(* PLC project Codesys Code Execution Speed Tests, CODESYS CODESYS V3.5 SP18 Patch 2, author Toni Kucic *)
(* stored: creationDateTime 2022-11-20T20:47:32.0555446, version 1.0, modificationDateTime 2022-11-20T20:38:51.788641, organization TK Automation *)
(* A collection of programs that measure various execution speeds of code. *)

TYPE dtTestStruct : STRUCT
  dummy1 : USINT := 255;
  Elem1 : INT := -1;
  Id : DWORD := 215215126;
  IdText : STRING := 'Testing for speed';
  dummy2 : ARRAY[0..11] OF DWORD;
  dummy4 : BOOL := FALSE;
  dummy5 : STRING(255) := 'Big array';
  dummy6 : LINT := 1211212723838939;
END_STRUCT;
END_TYPE

TYPE dtBitStruct : STRUCT
  bit1 : BIT;
  bit2 : BIT;
  bit3 : BIT;
  bit4 : BIT;
  bit5 : BIT;
  bit6 : BIT;
  bit7 : BIT;
  bit8 : BIT;
  bit9 : BIT;
  bit10 : BIT;
  bit11 : BIT;
  bit12 : BIT;
  bit13 : BIT;
  bit14 : BIT;
  bit15 : BIT;
  bit16 : BIT;
END_STRUCT;
END_TYPE

TYPE dtSpeedTest : STRUCT
  Results : ARRAY[0..9] OF LTIME;
  Desc : STRING(255);
  AverageExecTime : LTIME;
  OldTime : LTIME;
  ExecTime : LTIME;
END_STRUCT;
END_TYPE

PROGRAM x03_FloatingPointOperations
  VAR CONSTANT
    cNrRuns : USINT(0..9) := 5;
    cRepeatCalcTimes : UDINT := 1000000;  (* 1 Million times *)
  END_VAR
  VAR_INPUT
    vStart : BOOL := FALSE;
  END_VAR
  VAR
    vDone : BOOL := FALSE;
    vRunsCompleted : USINT := 0;
    vStartTime : LTIME;
    vTotalTime : LTIME;
    vTest1 : dtSpeedTest;
    vTest2 : dtSpeedTest;
    vTest3 : dtSpeedTest;
    vTest4 : dtSpeedTest;
    vTest5 : dtSpeedTest;
    vTest6 : dtSpeedTest;
    vTest7 : dtSpeedTest;
    vTest8 : dtSpeedTest;
    vTest9 : dtSpeedTest;
    i : UDINT;
    vInteger1 : INT := 1234;  (* Test vars *)
    vInteger2 : INT := 4231;
    vReal1 : REAL := 1234.4231;
    vReal2 : REAL := 4231.1234;
    vInteger3 : DINT := 1234;
    vInteger4 : DINT := 4231;
    vResult1 : INT;
    vResult2 : REAL;
    vResult3 : DINT;
    vResult4 : INT;
    vResult5 : REAL;
    vResult6 : DINT;
    vResult7 : INT;
    vResult8 : REAL;
    vResult9 : DINT;
  END_VAR

            (*Runs once on event's rising edge*)
vDone 		:= FALSE;
vStartTime 	:= LTIME();

FOR vRunsCompleted:=0 TO cNrRuns DO
	Measure();
END_FOR

vTotalTime := LTIME() - vStartTime;

vTest1.Desc				:= 'Time to add two integers 1 milion times';
vTest1.AverageExecTime 	:= calcAvg(vTest1.Results);
vTest2.Desc				:= 'Time to add two reals 1 milion times';
vTest2.AverageExecTime 	:= calcAvg(vTest2.Results);
vTest3.Desc				:= 'Time to add two DINTs (32b INT) 1 milion times';
vTest3.AverageExecTime 	:= calcAvg(vTest3.Results);
vTest4.Desc				:= 'Time to multiply two integers 1 milion times';
vTest4.AverageExecTime 	:= calcAvg(vTest4.Results);
vTest5.Desc				:= 'Time to multiply two reals 1 milion times';
vTest5.AverageExecTime 	:= calcAvg(vTest5.Results);
vTest6.Desc				:= 'Time to multiply two DINTs (32b INT) 1 milion times';
vTest6.AverageExecTime 	:= calcAvg(vTest6.Results);
vTest7.Desc				:= 'Time to divide two integers 1 milion times';
vTest7.AverageExecTime 	:= calcAvg(vTest7.Results);
vTest8.Desc				:= 'Time to divide two reals 1 milion times';
vTest8.AverageExecTime 	:= calcAvg(vTest8.Results);
vTest9.Desc				:= 'Time to divide two DINTs (32b INT) 1 milion times';
vTest9.AverageExecTime 	:= calcAvg(vTest9.Results);
	
vDone := TRUE;
vStart:= FALSE;

          

ACTION Measure:
                //------------CALCULATION A -------------------
vTest1.OldTime := LTIME();
FOR i:= 0 TO cRepeatCalcTimes DO
	vResult1 := vInteger1 + vInteger2;
END_FOR
vTest1.ExecTime := LTIME() - vTest1.OldTime;

//------------CALCULATION B -------------------
vTest2.OldTime := LTIME();
FOR i:= 0 TO cRepeatCalcTimes DO
	vResult2 := vReal1 + vReal2;
END_FOR
vTest2.ExecTime := LTIME() - vTest2.OldTime;

//------------CALCULATION C -------------------
vTest3.OldTime := LTIME();
FOR i:= 0 TO cRepeatCalcTimes DO
	vResult3 := vInteger3 + vInteger4;
END_FOR
vTest3.ExecTime := LTIME() - vTest3.OldTime;

//------------CALCULATION D -------------------
vTest4.OldTime := LTIME();
FOR i:= 0 TO cRepeatCalcTimes DO
	vResult4 := vInteger1 * vInteger2;
END_FOR
vTest4.ExecTime := LTIME() - vTest4.OldTime;

//------------CALCULATION E -------------------
vTest5.OldTime := LTIME();
FOR i:= 0 TO cRepeatCalcTimes DO
	vResult5 := vReal1 * vReal2;
END_FOR
vTest5.ExecTime := LTIME() - vTest5.OldTime;

//------------CALCULATION F -------------------
vTest6.OldTime := LTIME();
FOR i:= 0 TO cRepeatCalcTimes DO
	vResult6 := vInteger3 * vInteger4;
END_FOR
vTest6.ExecTime := LTIME() - vTest6.OldTime;

//------------CALCULATION G -------------------
vTest7.OldTime := LTIME();
FOR i:= 0 TO cRepeatCalcTimes DO
	vResult7 := vInteger1 / vInteger2;
END_FOR
vTest7.ExecTime := LTIME() - vTest7.OldTime;

//------------CALCULATION H -------------------
vTest8.OldTime := LTIME();
FOR i:= 0 TO cRepeatCalcTimes DO
	vResult8 := vReal1 / vReal2;
END_FOR
vTest8.ExecTime := LTIME() - vTest8.OldTime;

//------------CALCULATION I -------------------
vTest9.OldTime := LTIME();
FOR i:= 0 TO cRepeatCalcTimes DO
	vResult9 := vInteger3 / vInteger4;
END_FOR
vTest9.ExecTime := LTIME() - vTest9.OldTime;


//------------CATCH RESULTS---------------------
vTest1.Results[vRunsCompleted] := vTest1.ExecTime;
vTest2.Results[vRunsCompleted] := vTest2.ExecTime;
vTest3.Results[vRunsCompleted] := vTest3.ExecTime;
vTest4.Results[vRunsCompleted] := vTest4.ExecTime;
vTest5.Results[vRunsCompleted] := vTest5.ExecTime;
vTest6.Results[vRunsCompleted] := vTest6.ExecTime;
vTest7.Results[vRunsCompleted] := vTest7.ExecTime;
vTest8.Results[vRunsCompleted] := vTest8.ExecTime;
vTest9.Results[vRunsCompleted] := vTest9.ExecTime;
              
END_ACTION
END_PROGRAM

FUNCTION addTwoInts : INT
  VAR_IN_OUT
    int1 : INT;
    int2 : INT;
  END_VAR

            addTwoInts := int1 + int2;
          
END_FUNCTION

PROGRAM x04_FunctionOverhead
  VAR CONSTANT
    cNrRuns : USINT(0..9) := 5;
    cRepeatCalcTimes : UDINT := 1000000;  (* 1 Million times *)
  END_VAR
  VAR_INPUT
    vStart : BOOL := FALSE;
  END_VAR
  VAR
    vDone : BOOL := FALSE;
    vRunsCompleted : USINT := 0;
    vStartTime : LTIME;
    vTotalTime : LTIME;
    vTest1 : dtSpeedTest;
    vTest2 : dtSpeedTest;
    vTest3 : dtSpeedTest;
    i : UDINT;
    vInt1 : INT := 1;  (* Test vars *)
    vInt2 : INT := 2;
    vResult1 : INT;
    vResult2 : INT;
    vResult3 : INT;
  END_VAR

            (*Runs once on event's rising edge*)
vDone 		:= FALSE;
vStartTime 	:= LTIME();

FOR vRunsCompleted:=0 TO cNrRuns DO
	Measure();
END_FOR

vTotalTime := LTIME() - vStartTime;

vTest1.Desc				:= 'Calculation using just operands, 1 milion times';
vTest1.AverageExecTime 	:= calcAvg(vTest1.Results);
vTest2.Desc				:= 'Calculation using function, 1 milion times';
vTest2.AverageExecTime 	:= calcAvg(vTest2.Results);
vTest3.Desc				:= 'Calculation using PRG method, 1 milion times';
vTest3.AverageExecTime 	:= calcAvg(vTest3.Results);
	
vDone := TRUE;
vStart:= FALSE;

          

ACTION Measure:
                //------------CALCULATION A -------------------
vTest1.OldTime := LTIME();
FOR i:= 0 TO cRepeatCalcTimes DO
	vResult1 := vInt1 + vInt2;
END_FOR
vTest1.ExecTime := LTIME() - vTest1.OldTime;

//------------CALCULATION B -------------------
vTest2.OldTime := LTIME();
FOR i:= 0 TO cRepeatCalcTimes DO
	vResult2 := addTwoInts(vInt1, vInt2);
END_FOR
vTest2.ExecTime := LTIME() - vTest2.OldTime;

//------------CALCULATION C -------------------
vTest3.OldTime := LTIME();
FOR i:= 0 TO cRepeatCalcTimes DO
	vResult3 := addTwoNumbers(vInt1, vInt2);
END_FOR
vTest3.ExecTime := LTIME() - vTest3.OldTime;

//------------CATCH RESULTS---------------------
vTest1.Results[vRunsCompleted] := vTest1.ExecTime;
vTest2.Results[vRunsCompleted] := vTest2.ExecTime;
vTest3.Results[vRunsCompleted] := vTest3.ExecTime;
              
END_ACTION

METHOD addTwoNumbers : INT
  VAR_INPUT
    int1 : INT;
    int2 : INT;
  END_VAR
                  addTwoNumbers := int1 + int2;
                
END_METHOD
END_PROGRAM

PROGRAM x01_ImpactOfDynamicArrays
  VAR CONSTANT
    cNrRuns : USINT(0..9) := 5;
    cRepeatCalcTimes : UDINT := 1000000;  (* 1 Million times *)
  END_VAR
  VAR_INPUT
    vStart : BOOL := FALSE;
  END_VAR
  VAR
    vDone : BOOL := FALSE;
    vRunsCompleted : USINT := 0;
    vStartTime : LTIME;
    vTotalTime : LTIME;
    vTest1 : dtSpeedTest;
    vTest2 : dtSpeedTest;
    i : UDINT;
    vAvgTimeFun : LTIME;  (* Test vars *)
    vAvgTimeHardCoded : LTIME;
    vTimes : ARRAY[0..9] OF LTIME := [LTIME#1ms0us0ns, LTIME#2ms0us0ns, LTIME#3ms0us0ns, LTIME#4ms0us0ns, LTIME#5ms0us0ns, LTIME#6ms0us0ns, LTIME#7ms0us0ns, LTIME#8ms0us0ns, LTIME#9ms0us0ns, LTIME#10ms0us0ns];
    vTimes2 : ARRAY[0..9] OF LTIME := [LTIME#1ms0us0ns, LTIME#2ms0us0ns];
  END_VAR

            (*Runs once on event's rising edge*)
vDone 		:= FALSE;
vStartTime 	:= LTIME();

FOR vRunsCompleted:=0 TO cNrRuns DO
	Measure();
END_FOR

vTotalTime := LTIME() - vStartTime;

vTest1.Desc				:= 'Time took to run a function using ARRAY[*], 1 milion times';
vTest1.AverageExecTime  := calcAvg(vTest1.Results);

vTest2.Desc				:= 'Time took to run a function using fixed ARRAY[0..9], 1 milion times';
vTest2.AverageExecTime := calcAvg(vTest2.Results);

vDone := TRUE;
vStart:= FALSE;

          

ACTION Measure:
                //------------CALCULATION A -------------------
vTest1.OldTime := LTIME();
FOR i:= 0 TO cRepeatCalcTimes DO
	vAvgTimeFun := calcAvg(vTimes);
END_FOR
vTest1.ExecTime := LTIME() - vTest1.OldTime;

//------------CALCULATION B -------------------
vTest2.OldTime := LTIME();
FOR i:= 0 TO cRepeatCalcTimes DO
	vAvgTimeHardCoded := calcAvgFixed(vTimes2);
END_FOR
vTest2.ExecTime := LTIME() - vTest2.OldTime;

//------------CATCH RESULTS---------------------
vTest1.Results[vRunsCompleted] := vTest1.ExecTime;
vTest2.Results[vRunsCompleted] := vTest2.ExecTime;
              
END_ACTION
END_PROGRAM

PROGRAM x06_Combine2xByteToUint
  VAR CONSTANT
    cNrRuns : USINT(0..9) := 5;
    cRepeatCalcTimes : UDINT := 1000000;  (* 1 Million times *)
  END_VAR
  VAR_INPUT
    vStart : BOOL := FALSE;
  END_VAR
  VAR
    vDone : BOOL := FALSE;
    vRunsCompleted : USINT := 0;
    vStartTime : LTIME;
    vTotalTime : LTIME;
    vTest1 : dtSpeedTest;
    vTest2 : dtSpeedTest;
    vTest3 : dtSpeedTest;
    i : UDINT;
    vSHRInteger : UINT;  (* Test vars *)
    vMcpyInteger : UINT;
    vManualCpyInt : UINT;
    vBuffer : ARRAY[0..1] OF USINT := [16#55, 16#AA];
    vSHLOldTime : LTIME;
    vMcpyOldTime : LTIME;
    vSHLExecTime : LTIME;
    vMcpyExecTime : LTIME;
  END_VAR

            (*Runs once on event's rising edge*)
vDone 		:= FALSE;
vStartTime 	:= LTIME();

FOR vRunsCompleted:=0 TO cNrRuns DO
	Measure();
END_FOR

vTotalTime := LTIME() - vStartTime;

vTest1.Desc				:= 'Assembling an integer from two bytes (SHL), 1 milion times';
vTest1.AverageExecTime 	:= calcAvg(vTest1.Results);
vTest2.Desc				:= 'Assembling an integer from two bytes (SysMemCpy), 1 milion times';
vTest2.AverageExecTime 	:= calcAvg(vTest2.Results);
vTest3.Desc				:= 'Assembling an integer from two bytes by manually copying bits, 1 milion times';
vTest3.AverageExecTime 	:= calcAvg(vTest3.Results);
	
vDone := TRUE;
vStart:= FALSE;

          

ACTION Measure:
                //-------Assemble an UINT from two USINTs using SHL operator
vTest1.OldTime := LTIME();
FOR i:= 0 TO cRepeatCalcTimes DO
	vSHRInteger := vBuffer[0] + SHL(vBuffer[1],8);
END_FOR
vTest1.ExecTime := LTIME() - vTest1.OldTime;

//-------Assemble an UINT from two USINTs using MemCpy
vTest2.OldTime := LTIME();
FOR i:= 0 TO cRepeatCalcTimes DO
	SysMemCpy(ADR(vMcpyInteger), ADR(vBuffer) , SIZEOF(vMcpyInteger));
END_FOR
vTest2.ExecTime := LTIME() - vTest2.OldTime;

//-------Assemble an UINT from two USINTs by manually copying bits
vTest3.OldTime := LTIME();
FOR i:= 0 TO cRepeatCalcTimes DO
	vManualCpyInt.0 := vBuffer[0].0;
	vManualCpyInt.1 := vBuffer[0].1;
	vManualCpyInt.2 := vBuffer[0].2;
	vManualCpyInt.3 := vBuffer[0].3;
	vManualCpyInt.4 := vBuffer[0].4;
	vManualCpyInt.5 := vBuffer[0].5;
	vManualCpyInt.6 := vBuffer[0].6;
	vManualCpyInt.7 := vBuffer[0].7;
	
	vManualCpyInt.8 := vBuffer[1].0;
	vManualCpyInt.9 := vBuffer[1].1;
	vManualCpyInt.10 := vBuffer[1].2;
	vManualCpyInt.11 := vBuffer[1].3;
	vManualCpyInt.12 := vBuffer[1].4;
	vManualCpyInt.13 := vBuffer[1].5;
	vManualCpyInt.14 := vBuffer[1].6;
	vManualCpyInt.15 := vBuffer[1].7;

END_FOR
vTest3.ExecTime := LTIME() - vTest3.OldTime;

//Results
vTest1.Results[vRunsCompleted] := vTest1.ExecTime;
vTest2.Results[vRunsCompleted] := vTest2.ExecTime;
vTest3.Results[vRunsCompleted] := vTest3.ExecTime;
              
END_ACTION
END_PROGRAM

FUNCTION calcAVG : LTIME
  VAR_INPUT
    {attribute 'variable_length_array_original_scope' := 'Inout'}
    {attribute 'variable_length_array' := 'ARRAY[*] OF LTIME'}
    {attribute 'Dimensions' := '1'}
    Results : POINTER TO LTIME;
  END_VAR
  VAR
    i : DINT;
  END_VAR

            FOR i:=LOWER_BOUND(Results,1) TO UPPER_BOUND(Results,1) DO
	IF Results[i] = LTIME#0S THEN
		EXIT;
	END_IF
	calcAvg := calcAvg + Results[i];
END_FOR
calcAvg := calcAvg / MAX(1,i);
RETURN;
          
END_FUNCTION

PROGRAM x05_SysMemLib
  VAR CONSTANT
    cNrRuns : USINT(0..9) := 5;
    cRepeatCalcTimes : UDINT := 1000000;  (* 1 Million times *)
    cEmptyStruct : dtTestStruct;
  END_VAR
  VAR_INPUT
    vStart : BOOL := FALSE;
  END_VAR
  VAR
    vDone : BOOL := FALSE;
    vRunsCompleted : USINT := 0;
    vStartTime : LTIME;
    vTotalTime : LTIME;
    vTest1 : dtSpeedTest;
    vTest2 : dtSpeedTest;
    vTest3 : dtSpeedTest;
    vTest4 : dtSpeedTest;
    vTest5 : dtSpeedTest;
    vTest6 : dtSpeedTest;
    i : UDINT;
    vResultStruct1 : dtTestStruct;  (* Test variables *)
    vResultStruct2 : dtTestStruct;
    vResultStruct3 : dtTestStruct;
    vResultStruct4 : dtTestStruct;
    vResult5 : BOOL;
    vResult6 : BOOL;
  END_VAR

            (*Runs once on event's rising edge*)
vDone 		:= FALSE;
vStartTime 	:= LTIME();

FOR vRunsCompleted:=0 TO cNrRuns DO
	Measure();
END_FOR

vTotalTime := LTIME() - vStartTime;

vTest1.Desc				:= 'Setting a struct with an empty struct, 1 milion times';
vTest1.AverageExecTime 	:= calcAvg(vTest1.Results);
vTest2.Desc				:= 'Setting a struct with SysMemSet, 1 milion times';
vTest2.AverageExecTime 	:= calcAvg(vTest2.Results);
vTest3.Desc				:= 'Copy a struct to another struct, 1 milion times';
vTest3.AverageExecTime 	:= calcAvg(vTest3.Results);
vTest4.Desc				:= 'Copy a struct to another struct with memset, 1 milion times';
vTest4.AverageExecTime 	:= calcAvg(vTest4.Results);
vTest5.Desc				:= 'Compare a struct to another struct, 1 milion times';
vTest5.AverageExecTime 	:= calcAvg(vTest5.Results);
vTest6.Desc				:= 'Compare a struct to another struct with memcmp, 1 milion times';
vTest6.AverageExecTime 	:= calcAvg(vTest6.Results);
vDone := TRUE;
vStart:= FALSE;

          

ACTION Measure:
                //------------RESET STRUCT WITH A EMPTY STRUCT -------------------
vTest1.OldTime := LTIME();
FOR i:= 0 TO cRepeatCalcTimes DO
	vResultStruct1 := cEmptyStruct;
END_FOR
vTest1.ExecTime := LTIME() - vTest1.OldTime;

//------------RESET STRUCT WITH MEM SET -------------------
vTest2.OldTime := LTIME();
FOR i:= 0 TO cRepeatCalcTimes DO
	SysMemSet(ADR(vResultStruct2), 16#0 , SIZEOF(vResultStruct2));
END_FOR
vTest2.ExecTime := LTIME() - vTest2.OldTime;

//------------COPY STRUCT TO ANOTHER STRUCT -------------------
vTest3.OldTime := LTIME();
FOR i:= 0 TO cRepeatCalcTimes DO
	vResultStruct3 := cEmptyStruct;
END_FOR
vTest3.ExecTime := LTIME() - vTest3.OldTime;

//------------COPY STRUCT TO ANOTHER STRUCT MEMCPY -------------------
vTest4.OldTime := LTIME();
FOR i:= 0 TO cRepeatCalcTimes DO
	SysMemCpy(ADR(vResultStruct4), ADR(cEmptyStruct) , SIZEOF(cEmptyStruct));
END_FOR
vTest4.ExecTime := LTIME() - vTest4.OldTime;

//------------COMPARE STRUCT TO ANOTHER STRUCT -------------------
//NOTE: Codesys doesn't support complex struct comparing with = <>
vTest5.OldTime := LTIME();
FOR i:= 0 TO cRepeatCalcTimes DO
	vResult5 := vResultStruct3.dummy1 = cEmptyStruct.dummy1
			AND vResultStruct3.dummy2[0] = cEmptyStruct.dummy2[0]
			AND vResultStruct3.dummy2[1] = cEmptyStruct.dummy2[1]
			AND vResultStruct3.dummy2[2] = cEmptyStruct.dummy2[2]
			AND vResultStruct3.dummy2[3] = cEmptyStruct.dummy2[3]
			AND vResultStruct3.dummy2[4] = cEmptyStruct.dummy2[4]
			AND vResultStruct3.dummy2[5] = cEmptyStruct.dummy2[5]
			AND vResultStruct3.dummy2[6] = cEmptyStruct.dummy2[6]
			AND vResultStruct3.dummy2[7] = cEmptyStruct.dummy2[7]
			AND vResultStruct3.dummy2[8] = cEmptyStruct.dummy2[8]
			AND vResultStruct3.dummy2[9] = cEmptyStruct.dummy2[9]
			AND vResultStruct3.dummy2[10] = cEmptyStruct.dummy2[10]
			AND vResultStruct3.dummy2[11] = cEmptyStruct.dummy2[11]
			AND vResultStruct3.dummy4 = cEmptyStruct.dummy4
			AND vResultStruct3.dummy5 = cEmptyStruct.dummy5
			AND vResultStruct3.dummy6 = cEmptyStruct.dummy6
			AND vResultStruct3.Elem1 = cEmptyStruct.Elem1
			AND vResultStruct3.Id = cEmptyStruct.Id
			AND vResultStruct3.IdText = cEmptyStruct.IdText;
END_FOR
vTest5.ExecTime := LTIME() - vTest5.OldTime;

//------------COMPARE STRUCT TO ANOTHER STRUCT MEMCMP -------------------
vTest6.OldTime := LTIME();
FOR i:= 0 TO cRepeatCalcTimes DO
	vResult6 := SysMemCmp(ADR(vResultStruct4), ADR(cEmptyStruct),SIZEOF(cEmptyStruct)) = 0;
END_FOR
vTest6.ExecTime := LTIME() - vTest6.OldTime;

//------------CATCH RESULTS---------------------
vTest1.Results[vRunsCompleted] := vTest1.ExecTime;
vTest2.Results[vRunsCompleted] := vTest2.ExecTime;
vTest3.Results[vRunsCompleted] := vTest3.ExecTime;
vTest4.Results[vRunsCompleted] := vTest4.ExecTime;
vTest5.Results[vRunsCompleted] := vTest5.ExecTime;
vTest6.Results[vRunsCompleted] := vTest6.ExecTime;
              
END_ACTION
END_PROGRAM

PROGRAM x02_ExecSpeedOfLanguageTypes
  VAR CONSTANT
    cNrRuns : USINT(0..9) := 5;
    cRepeatCalcTimes : UDINT := 1000000;  (* 1 Million times *)
  END_VAR
  VAR_INPUT
    vStart : BOOL := FALSE;
  END_VAR
  VAR
    vDone : BOOL := FALSE;
    vRunsCompleted : USINT := 0;
    vStartTime : LTIME;
    vTotalTime : LTIME;
    vTest1 : dtSpeedTest;
    vTest2 : dtSpeedTest;
    vTest3 : dtSpeedTest;
    vTest4 : dtSpeedTest;
    i : UDINT;
    vInt1 : INT := 1;  (* Test vars *)
    vInt2 : INT := 2;
    vResult1 : INT;
    vResult2 : INT;
    vResult3 : INT;
    vResult4 : INT;
  END_VAR

            (*Runs once on event's rising edge*)
vDone 		:= FALSE;
vStartTime 	:= LTIME();

FOR vRunsCompleted:=0 TO cNrRuns DO
	Measure();
END_FOR

vTotalTime := LTIME() - vStartTime;

vTest1.Desc				:= 'Time function completed in LADDER, 1 milion times';
vTest1.AverageExecTime 	:= calcAvg(vTest1.Results);
vTest2.Desc				:= 'Time function completed in ST, 1 milion times';
vTest2.AverageExecTime 	:= calcAvg(vTest2.Results);
vTest3.Desc				:= 'Time function completed in FBD, 1 milion times';
vTest3.AverageExecTime 	:= calcAvg(vTest3.Results);
vTest4.Desc				:= 'Time function completed in CFC, 1 milion times';
vTest4.AverageExecTime 	:= calcAvg(vTest3.Results);

vDone := TRUE;
vStart:= FALSE;

          

ACTION Measure:
                //------------CALCULATION A -------------------
vTest1.OldTime := LTIME();
FOR i:= 0 TO cRepeatCalcTimes DO
	vResult1 := addTwoIntsLadder(vInt1, vInt2);
END_FOR
vTest1.ExecTime := LTIME() - vTest1.OldTime;

//------------CALCULATION B -------------------
vTest2.OldTime := LTIME();
FOR i:= 0 TO cRepeatCalcTimes DO
	vResult2 := addTwoIntsST(vInt1, vInt2);
END_FOR
vTest2.ExecTime := LTIME() - vTest2.OldTime;

//------------CALCULATION C -------------------
vTest3.OldTime := LTIME();
FOR i:= 0 TO cRepeatCalcTimes DO
	vResult3 := addTwoIntsFBD(vInt1, vInt2);
END_FOR
vTest3.ExecTime := LTIME() - vTest3.OldTime;

//------------CALCULATION D -------------------
vTest4.OldTime := LTIME();
FOR i:= 0 TO cRepeatCalcTimes DO
	vResult4 := addTwoIntsCFC(vInt1, vInt2);
END_FOR
vTest4.ExecTime := LTIME() - vTest4.OldTime;

//------------CATCH RESULTS---------------------
vTest1.Results[vRunsCompleted] := vTest1.ExecTime;
vTest2.Results[vRunsCompleted] := vTest2.ExecTime;
vTest3.Results[vRunsCompleted] := vTest3.ExecTime;
vTest4.Results[vRunsCompleted] := vTest4.ExecTime;
              
END_ACTION
END_PROGRAM

FUNCTION addTwoIntsLadder : INT
  VAR_INPUT
    Int1 : INT;
    Int2 : INT;
  END_VAR

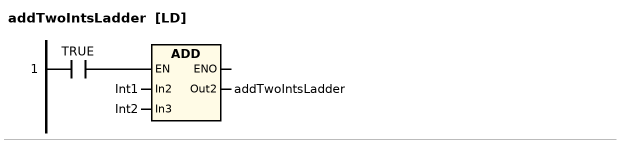
(* LD diagram, written out as Structured Text *)

IF TRUE THEN addTwoIntsLadder := Int1 + Int2; END_IF;
END_FUNCTION

FUNCTION addTwoIntsST : INT
  VAR_INPUT
    int1 : INT;
    int2 : INT;
  END_VAR

            addTwoIntsST := int1 + int2;
          
END_FUNCTION

FUNCTION addTwoIntsFBD : INT
  VAR_INPUT
    int1 : INT;
    int2 : INT;
  END_VAR

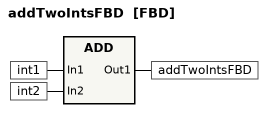
(* FBD diagram, written out as Structured Text *)
addTwoIntsFBD := int1 + int2;
END_FUNCTION

PROGRAM x07_StringOperations
  VAR CONSTANT
    cNrRuns : USINT(0..9) := 5;
    cRepeatCalcTimes : UDINT := 1000000;  (* 1 Million times *)
  END_VAR
  VAR_INPUT
    vStart : BOOL := FALSE;
  END_VAR
  VAR
    vDone : BOOL := FALSE;
    vRunsCompleted : USINT := 0;
    vStartTime : LTIME;
    vTotalTime : LTIME;
    vTest1 : dtSpeedTest;
    vTest2 : dtSpeedTest;
    vTest3 : dtSpeedTest;
    vTest4 : dtSpeedTest;
    vTest5 : dtSpeedTest;
    vTest6 : dtSpeedTest;
    i : UDINT;
    vString1 : STRING(255) := 'Test string1';  (* Test vars *)
    vString2 : STRING := 'Test string2';
    vString3 : STRING := 'a';
    vString4 : STRING := 'a';
    vByte : BYTE := 16#FF;
    vArrByte : ARRAY[0..255] OF BYTE;
    vResult1 : STRING(255);
    vResult2 : STRING;
    vResult3 : STRING;
    vResult4 : STRING(255);
    vResult5 : BYTE;
    vResult6 : ARRAY[0..255] OF BYTE;
    vSizes : ARRAY[0..3] OF UDINT;
  END_VAR

            (*Runs once on event's rising edge*)
vDone 		:= FALSE;

vSizes[0] := SIZEOF(vString1); //Size is 255 characters + zero char
vSizes[1] := SIZEOF(vString2); //Size is 80 characters + zero char, default if no size specified
vSizes[2] := SIZEOF(vResult3); //Size is 81, even though we concatenated 1 Million characters. The rest were chopped off
vSizes[3] := SIZEOF(vResult4); //Size is expected 256, other 744 characters chopped off

vStartTime 	:= LTIME();

FOR vRunsCompleted:=0 TO cNrRuns DO
	Measure();
END_FOR

vTotalTime := LTIME() - vStartTime;

vTest1.Desc				:= 'Time to copy a string[255] 1 Million times';
vTest1.AverageExecTime 	:= calcAvg(vTest1.Results);
vTest2.Desc				:= 'Time to copy a string 1 Million times';
vTest2.AverageExecTime 	:= calcAvg(vTest2.Results);
vTest3.Desc				:= 'Time to concatenate 1 Million times characters with STRING';
vTest3.AverageExecTime 	:= calcAvg(vTest3.Results);
vTest4.Desc				:= 'Time to concatenate 1 Million times  characters with STRING[255]';
vTest4.AverageExecTime 	:= calcAvg(vTest4.Results);
vTest5.Desc				:= 'Time to move a byte 1 Million times';
vTest5.AverageExecTime 	:= calcAvg(vTest5.Results);
vTest6.Desc				:= 'Time to copy an array of 255 BYTE 1 Million times';
vTest6.AverageExecTime 	:= calcAvg(vTest6.Results);
	
vDone := TRUE;
vStart:= FALSE;

          

ACTION Measure:
                //------------CALCULATION A -------------------
vTest1.OldTime := LTIME();
FOR i:= 0 TO cRepeatCalcTimes DO
	vResult1 := vString1;
END_FOR
vTest1.ExecTime := LTIME() - vTest1.OldTime;

//------------CALCULATION B -------------------
vTest2.OldTime := LTIME();
FOR i:= 0 TO cRepeatCalcTimes DO
	vResult2 := vString2;
END_FOR
vTest2.ExecTime := LTIME() - vTest2.OldTime;

//------------CALCULATION C -------------------
vTest3.OldTime := LTIME();
FOR i:= 0 TO cRepeatCalcTimes DO
	vResult3 := CONCAT(vResult3, vString3);
END_FOR
vTest3.ExecTime := LTIME() - vTest3.OldTime;

//------------CALCULATION D -------------------
vTest4.OldTime := LTIME();
FOR i:= 0 TO cRepeatCalcTimes DO
	vResult4 := CONCAT(vResult4, vString4);
END_FOR
vTest4.ExecTime := LTIME() - vTest4.OldTime;

//------------CALCULATION E -------------------
vTest5.OldTime := LTIME();
FOR i:= 0 TO cRepeatCalcTimes DO
	vResult5 := vByte;
END_FOR
vTest5.ExecTime := LTIME() - vTest5.OldTime;

//------------CALCULATION F -------------------
vTest6.OldTime := LTIME();
FOR i:= 0 TO cRepeatCalcTimes DO
	vResult6 := vArrByte;
END_FOR
vTest6.ExecTime := LTIME() - vTest6.OldTime;

//------------CATCH RESULTS---------------------
vTest1.Results[vRunsCompleted] := vTest1.ExecTime;
vTest2.Results[vRunsCompleted] := vTest2.ExecTime;
vTest3.Results[vRunsCompleted] := vTest3.ExecTime;
vTest4.Results[vRunsCompleted] := vTest4.ExecTime;
vTest5.Results[vRunsCompleted] := vTest5.ExecTime;
vTest6.Results[vRunsCompleted] := vTest6.ExecTime;
              
END_ACTION
END_PROGRAM

PROGRAM x08_CheckingBools
  VAR CONSTANT
    cNrRuns : USINT(0..9) := 5;
    cRepeatCalcTimes : UDINT := 1000000;  (* 1 Million times *)
  END_VAR
  VAR_INPUT
    vStart : BOOL := FALSE;
  END_VAR
  VAR
    vDone : BOOL := FALSE;
    vRunsCompleted : USINT := 0;
    vStartTime : LTIME;
    vTotalTime : LTIME;
    vTest1 : dtSpeedTest;
    vTest2 : dtSpeedTest;
    vTest3 : dtSpeedTest;
    vTest4 : dtSpeedTest;
    vTest5 : dtSpeedTest;
    i : UDINT;
    vBool : BOOL := TRUE;  (* Test vars *)
    vResult : BOOL;
    vCounter : UINT := 0;
    vCastedUint : UINT;
  END_VAR

            (*Runs once on event's rising edge*)
vDone 		:= FALSE;
vStartTime 	:= LTIME();

FOR vRunsCompleted:=0 TO cNrRuns DO
	Measure();
END_FOR

vTotalTime := LTIME() - vStartTime;

vTest1.Desc				:= 'Time to run IF vBool = TRUE THEN 1 Million times';
vTest1.AverageExecTime 	:= calcAvg(vTest1.Results);
vTest2.Desc				:= 'Time to run IF vBool THEN 1 Million times';
vTest2.AverageExecTime 	:= calcAvg(vTest2.Results);
vTest3.Desc				:= 'Time to increment a counter using if sentence 1 Million times';
vTest3.AverageExecTime 	:= calcAvg(vTest3.Results);
vTest4.Desc				:= 'Time to increment a counter using bool to UINT 1 Million times';
vTest4.AverageExecTime 	:= calcAvg(vTest4.Results);
vTest5.Desc				:= 'Time to cast a bool to UINT 1 Million times';
vTest5.AverageExecTime 	:= calcAvg(vTest5.Results);
	
vDone := TRUE;
vStart:= FALSE;

          

ACTION Measure:
                //------------CALCULATION A -------------------
vTest1.OldTime := LTIME();
FOR i:= 0 TO cRepeatCalcTimes DO
	IF vBool = TRUE THEN
		vResult := vBool;
	END_IF
END_FOR
vTest1.ExecTime := LTIME() - vTest1.OldTime;

//------------CALCULATION B -------------------
vTest2.OldTime := LTIME();
FOR i:= 0 TO cRepeatCalcTimes DO
	IF vBool THEN
		vResult := vBool;
	END_IF
END_FOR
vTest2.ExecTime := LTIME() - vTest2.OldTime;

//------------CALCULATION C -------------------
vTest3.OldTime := LTIME();
FOR i:= 0 TO cRepeatCalcTimes DO
	IF vBool THEN
		vCounter := vCounter + 1;
	END_IF
END_FOR
vTest3.ExecTime := LTIME() - vTest3.OldTime;

//------------CALCULATION D -------------------
vTest4.OldTime := LTIME();
FOR i:= 0 TO cRepeatCalcTimes DO
	vCounter := vCounter + BOOL_TO_UINT(vBool);
END_FOR
vTest4.ExecTime := LTIME() - vTest4.OldTime;

//------------CALCULATION D -------------------
vTest5.OldTime := LTIME();
FOR i:= 0 TO cRepeatCalcTimes DO
	vCastedUint := BOOL_TO_UINT(vBool);
END_FOR
vTest5.ExecTime := LTIME() - vTest5.OldTime;

//------------CATCH RESULTS---------------------
vTest1.Results[vRunsCompleted] := vTest1.ExecTime;
vTest2.Results[vRunsCompleted] := vTest2.ExecTime;
vTest3.Results[vRunsCompleted] := vTest3.ExecTime;
vTest4.Results[vRunsCompleted] := vTest4.ExecTime;
vTest5.Results[vRunsCompleted] := vTest5.ExecTime;
              
END_ACTION
END_PROGRAM

PROGRAM x09_CaseVsIfElsif
  VAR CONSTANT
    cNrRuns : USINT(0..9) := 5;
    cRepeatCalcTimes : UDINT := 1000000;  (* 1 Million times *)
  END_VAR
  VAR_INPUT
    vStart : BOOL := FALSE;
  END_VAR
  VAR
    vDone : BOOL := FALSE;
    vRunsCompleted : USINT := 0;
    vStartTime : LTIME;
    vTotalTime : LTIME;
    vTest1 : dtSpeedTest;
    vTest2 : dtSpeedTest;
    vTest3 : dtSpeedTest;
    vTest4 : dtSpeedTest;
    vTest5 : dtSpeedTest;
    vTest6 : dtSpeedTest;
    i : UDINT;
    vFirstIndex : INT := 15;  (* Test vars *)
    vMiddleIndex : INT := 50;
    vLastIndex : INT := 99;
    vResultFirst : INT;  (* Should be 0 *)
    vResultMiddle : INT;  (* Should be 50 *)
    vResultLast : INT;  (* Should be 99 *)
  END_VAR

            (*Runs once on event's rising edge*)
vDone 		:= FALSE;
vStartTime 	:= LTIME();

FOR vRunsCompleted:=0 TO cNrRuns DO
	Measure();
END_FOR

vTotalTime := LTIME() - vStartTime;

vTest1.Desc				:= 'Time to run first branch of IF ELSIF 1 Million times';
vTest1.AverageExecTime 	:= calcAvg(vTest1.Results);
vTest2.Desc				:= 'Time to run middle branch of IF ELSIF 1 Million times';
vTest2.AverageExecTime 	:= calcAvg(vTest2.Results);
vTest3.Desc				:= 'Time to run last branch of IF ELSIF 1 Million times';
vTest3.AverageExecTime 	:= calcAvg(vTest3.Results);
vTest4.Desc				:= 'Time to run first branch of CASE 1 Million times';
vTest4.AverageExecTime 	:= calcAvg(vTest4.Results);
vTest5.Desc				:= 'Time to run middle branch of CASE 1 Million times';
vTest5.AverageExecTime 	:= calcAvg(vTest5.Results);
vTest6.Desc				:= 'Time to run last branch of CASE 1 Million times';
vTest6.AverageExecTime 	:= calcAvg(vTest6.Results);
	
vDone := TRUE;
vStart:= FALSE;

          

ACTION Measure:
                //------------CALCULATION A -------------------
vTest1.OldTime := LTIME();
FOR i:= 0 TO cRepeatCalcTimes DO
	vResultFirst := returnIndexIfElsif(vFirstIndex);
END_FOR
vTest1.ExecTime := LTIME() - vTest1.OldTime;

//------------CALCULATION B -------------------
vTest2.OldTime := LTIME();
FOR i:= 0 TO cRepeatCalcTimes DO
	vResultMiddle := returnIndexIfElsif(vMiddleIndex);
END_FOR
vTest2.ExecTime := LTIME() - vTest2.OldTime;

//------------CALCULATION C -------------------
vTest3.OldTime := LTIME();
FOR i:= 0 TO cRepeatCalcTimes DO
	vResultLast := returnIndexIfElsif(vLastIndex);
END_FOR
vTest3.ExecTime := LTIME() - vTest3.OldTime;

//------------CALCULATION D -------------------
vTest4.OldTime := LTIME();
FOR i:= 0 TO cRepeatCalcTimes DO
	vResultFirst := returnIndexCase(vFirstIndex);
END_FOR
vTest4.ExecTime := LTIME() - vTest4.OldTime;

//------------CALCULATION E -------------------
vTest5.OldTime := LTIME();
FOR i:= 0 TO cRepeatCalcTimes DO
	vResultMiddle := returnIndexCase(vMiddleIndex);
END_FOR
vTest5.ExecTime := LTIME() - vTest5.OldTime;

//------------CALCULATION F -------------------
vTest6.OldTime := LTIME();
FOR i:= 0 TO cRepeatCalcTimes DO
	vResultLast := returnIndexCase(vLastIndex);
END_FOR
vTest6.ExecTime := LTIME() - vTest6.OldTime;

//------------CATCH RESULTS---------------------
vTest1.Results[vRunsCompleted] := vTest1.ExecTime;
vTest2.Results[vRunsCompleted] := vTest2.ExecTime;
vTest3.Results[vRunsCompleted] := vTest3.ExecTime;
vTest4.Results[vRunsCompleted] := vTest4.ExecTime;
vTest5.Results[vRunsCompleted] := vTest5.ExecTime;
vTest6.Results[vRunsCompleted] := vTest6.ExecTime;
              
END_ACTION

METHOD returnIndexIfElsif : INT
  VAR_INPUT
    searchValue : INT;
  END_VAR
                  IF searchValue = 0 THEN
        returnIndexIfElsif:=0;
        RETURN;

ELSIF searchValue = 1 THEN
        returnIndexIfElsif:= 1;
        RETURN;

ELSIF searchValue = 2 THEN
        returnIndexIfElsif:= 2;
        RETURN;

ELSIF searchValue = 3 THEN
        returnIndexIfElsif:= 3;
        RETURN;

ELSIF searchValue = 4 THEN
        returnIndexIfElsif:= 4;
        RETURN;

ELSIF searchValue = 5 THEN
        returnIndexIfElsif:= 5;
        RETURN;

ELSIF searchValue = 6 THEN
        returnIndexIfElsif:= 6;
        RETURN;

ELSIF searchValue = 7 THEN
        returnIndexIfElsif:= 7;
        RETURN;

ELSIF searchValue = 8 THEN
        returnIndexIfElsif:= 8;
        RETURN;

ELSIF searchValue = 9 THEN
        returnIndexIfElsif:= 9;
        RETURN;

ELSIF searchValue = 10 THEN
        returnIndexIfElsif:= 10;
        RETURN;

ELSIF searchValue = 11 THEN
        returnIndexIfElsif:= 11;
        RETURN;

ELSIF searchValue = 12 THEN
        returnIndexIfElsif:= 12;
        RETURN;

ELSIF searchValue = 13 THEN
        returnIndexIfElsif:= 13;
        RETURN;

ELSIF searchValue = 14 THEN
        returnIndexIfElsif:= 14;
        RETURN;

ELSIF searchValue = 15 THEN
        returnIndexIfElsif:= 15;
        RETURN;

ELSIF searchValue = 16 THEN
        returnIndexIfElsif:= 16;
        RETURN;

ELSIF searchValue = 17 THEN
        returnIndexIfElsif:= 17;
        RETURN;

ELSIF searchValue = 18 THEN
        returnIndexIfElsif:= 18;
        RETURN;

ELSIF searchValue = 19 THEN
        returnIndexIfElsif:= 19;
        RETURN;

ELSIF searchValue = 20 THEN
        returnIndexIfElsif:= 20;
        RETURN;

ELSIF searchValue = 21 THEN
        returnIndexIfElsif:= 21;
        RETURN;

ELSIF searchValue = 22 THEN
        returnIndexIfElsif:= 22;
        RETURN;

ELSIF searchValue = 23 THEN
        returnIndexIfElsif:= 23;
        RETURN;

ELSIF searchValue = 24 THEN
        returnIndexIfElsif:= 24;
        RETURN;

ELSIF searchValue = 25 THEN
        returnIndexIfElsif:= 25;
        RETURN;

ELSIF searchValue = 26 THEN
        returnIndexIfElsif:= 26;
        RETURN;

ELSIF searchValue = 27 THEN
        returnIndexIfElsif:= 27;
        RETURN;

ELSIF searchValue = 28 THEN
        returnIndexIfElsif:= 28;
        RETURN;

ELSIF searchValue = 29 THEN
        returnIndexIfElsif:= 29;
        RETURN;

ELSIF searchValue = 30 THEN
        returnIndexIfElsif:= 30;
        RETURN;

ELSIF searchValue = 31 THEN
        returnIndexIfElsif:= 31;
        RETURN;

ELSIF searchValue = 32 THEN
        returnIndexIfElsif:= 32;
        RETURN;

ELSIF searchValue = 33 THEN
        returnIndexIfElsif:= 33;
        RETURN;

ELSIF searchValue = 34 THEN
        returnIndexIfElsif:= 34;
        RETURN;

ELSIF searchValue = 35 THEN
        returnIndexIfElsif:= 35;
        RETURN;

ELSIF searchValue = 36 THEN
        returnIndexIfElsif:= 36;
        RETURN;

ELSIF searchValue = 37 THEN
        returnIndexIfElsif:= 37;
        RETURN;

ELSIF searchValue = 38 THEN
        returnIndexIfElsif:= 38;
        RETURN;

ELSIF searchValue = 39 THEN
        returnIndexIfElsif:= 39;
        RETURN;

ELSIF searchValue = 40 THEN
        returnIndexIfElsif:= 40;
        RETURN;

ELSIF searchValue = 41 THEN
        returnIndexIfElsif:= 41;
        RETURN;

ELSIF searchValue = 42 THEN
        returnIndexIfElsif:= 42;
        RETURN;

ELSIF searchValue = 43 THEN
        returnIndexIfElsif:= 43;
        RETURN;

ELSIF searchValue = 44 THEN
        returnIndexIfElsif:= 44;
        RETURN;

ELSIF searchValue = 45 THEN
        returnIndexIfElsif:= 45;
        RETURN;

ELSIF searchValue = 46 THEN
        returnIndexIfElsif:= 46;
        RETURN;

ELSIF searchValue = 47 THEN
        returnIndexIfElsif:= 47;
        RETURN;

ELSIF searchValue = 48 THEN
        returnIndexIfElsif:= 48;
        RETURN;

ELSIF searchValue = 49 THEN
        returnIndexIfElsif:= 49;
        RETURN;

ELSIF searchValue = 50 THEN
        returnIndexIfElsif:= 50;
        RETURN;

ELSIF searchValue = 51 THEN
        returnIndexIfElsif:= 51;
        RETURN;

ELSIF searchValue = 52 THEN
        returnIndexIfElsif:= 52;
        RETURN;

ELSIF searchValue = 53 THEN
        returnIndexIfElsif:= 53;
        RETURN;

ELSIF searchValue = 54 THEN
        returnIndexIfElsif:= 54;
        RETURN;

ELSIF searchValue = 55 THEN
        returnIndexIfElsif:= 55;
        RETURN;

ELSIF searchValue = 56 THEN
        returnIndexIfElsif:= 56;
        RETURN;

ELSIF searchValue = 57 THEN
        returnIndexIfElsif:= 57;
        RETURN;

ELSIF searchValue = 58 THEN
        returnIndexIfElsif:= 58;
        RETURN;

ELSIF searchValue = 59 THEN
        returnIndexIfElsif:= 59;
        RETURN;

ELSIF searchValue = 60 THEN
        returnIndexIfElsif:= 60;
        RETURN;

ELSIF searchValue = 61 THEN
        returnIndexIfElsif:= 61;
        RETURN;

ELSIF searchValue = 62 THEN
        returnIndexIfElsif:= 62;
        RETURN;

ELSIF searchValue = 63 THEN
        returnIndexIfElsif:= 63;
        RETURN;

ELSIF searchValue = 64 THEN
        returnIndexIfElsif:= 64;
        RETURN;

ELSIF searchValue = 65 THEN
        returnIndexIfElsif:= 65;
        RETURN;

ELSIF searchValue = 66 THEN
        returnIndexIfElsif:= 66;
        RETURN;

ELSIF searchValue = 67 THEN
        returnIndexIfElsif:= 67;
        RETURN;

ELSIF searchValue = 68 THEN
        returnIndexIfElsif:= 68;
        RETURN;

ELSIF searchValue = 69 THEN
        returnIndexIfElsif:= 69;
        RETURN;

ELSIF searchValue = 70 THEN
        returnIndexIfElsif:= 70;
        RETURN;

ELSIF searchValue = 71 THEN
        returnIndexIfElsif:= 71;
        RETURN;

ELSIF searchValue = 72 THEN
        returnIndexIfElsif:= 72;
        RETURN;

ELSIF searchValue = 73 THEN
        returnIndexIfElsif:= 73;
        RETURN;

ELSIF searchValue = 74 THEN
        returnIndexIfElsif:= 74;
        RETURN;

ELSIF searchValue = 75 THEN
        returnIndexIfElsif:= 75;
        RETURN;

ELSIF searchValue = 76 THEN
        returnIndexIfElsif:= 76;
        RETURN;

ELSIF searchValue = 77 THEN
        returnIndexIfElsif:= 77;
        RETURN;

ELSIF searchValue = 78 THEN
        returnIndexIfElsif:= 78;
        RETURN;

ELSIF searchValue = 79 THEN
        returnIndexIfElsif:= 79;
        RETURN;

ELSIF searchValue = 80 THEN
        returnIndexIfElsif:= 80;
        RETURN;

ELSIF searchValue = 81 THEN
        returnIndexIfElsif:= 81;
        RETURN;

ELSIF searchValue = 82 THEN
        returnIndexIfElsif:= 82;
        RETURN;

ELSIF searchValue = 83 THEN
        returnIndexIfElsif:= 83;
        RETURN;

ELSIF searchValue = 84 THEN
        returnIndexIfElsif:= 84;
        RETURN;

ELSIF searchValue = 85 THEN
        returnIndexIfElsif:= 85;
        RETURN;

ELSIF searchValue = 86 THEN
        returnIndexIfElsif:= 86;
        RETURN;

ELSIF searchValue = 87 THEN
        returnIndexIfElsif:= 87;
        RETURN;

ELSIF searchValue = 88 THEN
        returnIndexIfElsif:= 88;
        RETURN;

ELSIF searchValue = 89 THEN
        returnIndexIfElsif:= 89;
        RETURN;

ELSIF searchValue = 90 THEN
        returnIndexIfElsif:= 90;
        RETURN;

ELSIF searchValue = 91 THEN
        returnIndexIfElsif:= 91;
        RETURN;

ELSIF searchValue = 92 THEN
        returnIndexIfElsif:= 92;
        RETURN;

ELSIF searchValue = 93 THEN
        returnIndexIfElsif:= 93;
        RETURN;

ELSIF searchValue = 94 THEN
        returnIndexIfElsif:= 94;
        RETURN;

ELSIF searchValue = 95 THEN
        returnIndexIfElsif:= 95;
        RETURN;

ELSIF searchValue = 96 THEN
        returnIndexIfElsif:= 96;
        RETURN;

ELSIF searchValue = 97 THEN
        returnIndexIfElsif:= 97;
        RETURN;

ELSIF searchValue = 98 THEN
        returnIndexIfElsif:= 98;
        RETURN;

ELSIF searchValue = 99 THEN
        returnIndexIfElsif:= 99;
        RETURN;

END_IF
                
END_METHOD

METHOD returnIndexCase : INT
  VAR_INPUT
    searchValue : INT;
  END_VAR
                  CASE searchValue OF

        0: returnIndexCase := 0;
        RETURN;

        1: returnIndexCase := 1;
        RETURN;

        2: returnIndexCase := 2;
        RETURN;

        3: returnIndexCase := 3;
        RETURN;

        4: returnIndexCase := 4;
        RETURN;

        5: returnIndexCase := 5;
        RETURN;

        6: returnIndexCase := 6;
        RETURN;

        7: returnIndexCase := 7;
        RETURN;

        8: returnIndexCase := 8;
        RETURN;

        9: returnIndexCase := 9;
        RETURN;

        10: returnIndexCase := 10;
        RETURN;

        11: returnIndexCase := 11;
        RETURN;

        12: returnIndexCase := 12;
        RETURN;

        13: returnIndexCase := 13;
        RETURN;

        14: returnIndexCase := 14;
        RETURN;

        15: returnIndexCase := 15;
        RETURN;

        16: returnIndexCase := 16;
        RETURN;

        17: returnIndexCase := 17;
        RETURN;

        18: returnIndexCase := 18;
        RETURN;

        19: returnIndexCase := 19;
        RETURN;

        20: returnIndexCase := 20;
        RETURN;

        21: returnIndexCase := 21;
        RETURN;

        22: returnIndexCase := 22;
        RETURN;

        23: returnIndexCase := 23;
        RETURN;

        24: returnIndexCase := 24;
        RETURN;

        25: returnIndexCase := 25;
        RETURN;

        26: returnIndexCase := 26;
        RETURN;

        27: returnIndexCase := 27;
        RETURN;

        28: returnIndexCase := 28;
        RETURN;

        29: returnIndexCase := 29;
        RETURN;

        30: returnIndexCase := 30;
        RETURN;

        31: returnIndexCase := 31;
        RETURN;

        32: returnIndexCase := 32;
        RETURN;

        33: returnIndexCase := 33;
        RETURN;

        34: returnIndexCase := 34;
        RETURN;

        35: returnIndexCase := 35;
        RETURN;

        36: returnIndexCase := 36;
        RETURN;

        37: returnIndexCase := 37;
        RETURN;

        38: returnIndexCase := 38;
        RETURN;

        39: returnIndexCase := 39;
        RETURN;

        40: returnIndexCase := 40;
        RETURN;

        41: returnIndexCase := 41;
        RETURN;

        42: returnIndexCase := 42;
        RETURN;

        43: returnIndexCase := 43;
        RETURN;

        44: returnIndexCase := 44;
        RETURN;

        45: returnIndexCase := 45;
        RETURN;

        46: returnIndexCase := 46;
        RETURN;

        47: returnIndexCase := 47;
        RETURN;

        48: returnIndexCase := 48;
        RETURN;

        49: returnIndexCase := 49;
        RETURN;

        50: returnIndexCase := 50;
        RETURN;

        51: returnIndexCase := 51;
        RETURN;

        52: returnIndexCase := 52;
        RETURN;

        53: returnIndexCase := 53;
        RETURN;

        54: returnIndexCase := 54;
        RETURN;

        55: returnIndexCase := 55;
        RETURN;

        56: returnIndexCase := 56;
        RETURN;

        57: returnIndexCase := 57;
        RETURN;

        58: returnIndexCase := 58;
        RETURN;

        59: returnIndexCase := 59;
        RETURN;

        60: returnIndexCase := 60;
        RETURN;

        61: returnIndexCase := 61;
        RETURN;

        62: returnIndexCase := 62;
        RETURN;

        63: returnIndexCase := 63;
        RETURN;

        64: returnIndexCase := 64;
        RETURN;

        65: returnIndexCase := 65;
        RETURN;

        66: returnIndexCase := 66;
        RETURN;

        67: returnIndexCase := 67;
        RETURN;

        68: returnIndexCase := 68;
        RETURN;

        69: returnIndexCase := 69;
        RETURN;

        70: returnIndexCase := 70;
        RETURN;

        71: returnIndexCase := 71;
        RETURN;

        72: returnIndexCase := 72;
        RETURN;

        73: returnIndexCase := 73;
        RETURN;

        74: returnIndexCase := 74;
        RETURN;

        75: returnIndexCase := 75;
        RETURN;

        76: returnIndexCase := 76;
        RETURN;

        77: returnIndexCase := 77;
        RETURN;

        78: returnIndexCase := 78;
        RETURN;

        79: returnIndexCase := 79;
        RETURN;

        80: returnIndexCase := 80;
        RETURN;

        81: returnIndexCase := 81;
        RETURN;

        82: returnIndexCase := 82;
        RETURN;

        83: returnIndexCase := 83;
        RETURN;

        84: returnIndexCase := 84;
        RETURN;

        85: returnIndexCase := 85;
        RETURN;

        86: returnIndexCase := 86;
        RETURN;

        87: returnIndexCase := 87;
        RETURN;

        88: returnIndexCase := 88;
        RETURN;

        89: returnIndexCase := 89;
        RETURN;

        90: returnIndexCase := 90;
        RETURN;

        91: returnIndexCase := 91;
        RETURN;

        92: returnIndexCase := 92;
        RETURN;

        93: returnIndexCase := 93;
        RETURN;

        94: returnIndexCase := 94;
        RETURN;

        95: returnIndexCase := 95;
        RETURN;

        96: returnIndexCase := 96;
        RETURN;

        97: returnIndexCase := 97;
        RETURN;

        98: returnIndexCase := 98;
        RETURN;

        99: returnIndexCase := 99;
        RETURN;

END_CASE
                
END_METHOD
END_PROGRAM

PROGRAM x10_1_BitAccess
  VAR CONSTANT
    cNrRuns : USINT(0..9) := 5;
    cRepeatCalcTimes : UDINT := 1000000;  (* 1 Million times *)
  END_VAR
  VAR_INPUT
    vStart : BOOL := FALSE;
  END_VAR
  VAR
    vDone : BOOL := FALSE;
    vRunsCompleted : USINT := 0;
    vStartTime : LTIME;
    vTotalTime : LTIME;
    vTest1 : dtSpeedTest;
    vTest2 : dtSpeedTest;
    vTest3 : dtSpeedTest;
    i : UDINT;
    vCodesysBits : dtBitStruct;  (* Test vars *)
    vNormalInt : UINT := 16#5555;
    vResult1 : BOOL;
    vResult2 : BOOL;
    vResult3 : BOOL;
  END_VAR

            (*Runs once on event's rising edge*)
vDone 		:= FALSE;
vStartTime 	:= LTIME();

FOR vRunsCompleted:=0 TO cNrRuns DO
	Measure();
END_FOR

vTotalTime := LTIME() - vStartTime;

vTest1.Desc				:= 'Time to access bit 3 1 Million times in codesys bit struct';
vTest1.AverageExecTime 	:= calcAvg(vTest1.Results);
vTest2.Desc				:= 'Time to access bit 3 1 Million times in normal integer using . notation';
vTest2.AverageExecTime 	:= calcAvg(vTest2.Results);
vTest3.Desc				:= 'Time to access bit 3 1 Million times in normal integer using bit masking';
vTest3.AverageExecTime 	:= calcAvg(vTest3.Results);
	
vDone := TRUE;
vStart:= FALSE;

          

ACTION Measure:
                //------------CALCULATION A -------------------
vTest1.OldTime := LTIME();
FOR i:= 0 TO cRepeatCalcTimes DO
	vResult1 := checkBit_bitStruct(vCodesysBits,2);
END_FOR
vTest1.ExecTime := LTIME() - vTest1.OldTime;

//------------CALCULATION B -------------------
vTest2.OldTime := LTIME();
FOR i:= 0 TO cRepeatCalcTimes DO
	vResult2 := checkBit_dotNot(vNormalInt,2);
END_FOR
vTest2.ExecTime := LTIME() - vTest2.OldTime;

//------------CALCULATION C -------------------
vTest3.OldTime := LTIME();
FOR i:= 0 TO cRepeatCalcTimes DO
	vResult3 := checkBit_bitmask(vNormalInt, 2);
END_FOR
vTest3.ExecTime := LTIME() - vTest3.OldTime;

//------------CATCH RESULTS---------------------
vTest1.Results[vRunsCompleted] := vTest1.ExecTime;
vTest2.Results[vRunsCompleted] := vTest2.ExecTime;
vTest3.Results[vRunsCompleted] := vTest3.ExecTime;
              
END_ACTION
END_PROGRAM

PROGRAM x10_3_BitMath
  VAR CONSTANT
    cNrRuns : USINT(0..9) := 5;
    cRepeatCalcTimes : UDINT := 1000000;  (* 1 Million times *)
  END_VAR
  VAR_INPUT
    vStart : BOOL := FALSE;
  END_VAR
  VAR
    vDone : BOOL := FALSE;
    vRunsCompleted : USINT := 0;
    vStartTime : LTIME;
    vTotalTime : LTIME;
    vTest1 : dtSpeedTest;
    vTest2 : dtSpeedTest;
    vTest3 : dtSpeedTest;
    i : UDINT;
    vCodesysBits : dtBitStruct := (bit1 := TRUE, bit2 := TRUE, bit3 := FALSE);  (* Test vars *)
    vNormalInt : UINT := 2#11;
    vNormalInt2 : UINT := 2#11;
    vNormalInt3 : UINT := 2#11;
  END_VAR

            (*Runs once on event's rising edge*)
vDone 		:= FALSE;
vStartTime 	:= LTIME();

FOR vRunsCompleted:=0 TO cNrRuns DO
	Measure();
END_FOR

vTotalTime := LTIME() - vStartTime;

vTest1.Desc				:= 'Time to and two bits and save it to another bit 1 Million times using codesys bit struct';
vTest1.AverageExecTime 	:= calcAvg(vTest1.Results);
vTest2.Desc				:= 'Time to and two bits and save it to another bit 1 Million times using . notation';
vTest2.AverageExecTime 	:= calcAvg(vTest2.Results);
vTest3.Desc				:= 'Time to and two bits and save it to another bit 1 Million times using bit masking';
vTest3.AverageExecTime 	:= calcAvg(vTest3.Results);
	
vDone := TRUE;
vStart:= FALSE;

          

ACTION Measure:
                //------------CALCULATION A -------------------
vTest1.OldTime := LTIME();
FOR i:= 0 TO cRepeatCalcTimes DO
	setBitToValue_bitStruct(vCodesysBits, 2, checkBit_bitStruct(vCodesysBits, 0) AND checkBit_bitStruct(vCodesysBits, 1));
END_FOR
vTest1.ExecTime := LTIME() - vTest1.OldTime;

//------------CALCULATION B -------------------
vTest2.OldTime := LTIME();
FOR i:= 0 TO cRepeatCalcTimes DO
	setBitToValue_dotNot(vNormalInt, 2, checkBit_dotNot(vNormalInt, 0) AND checkBit_dotNot(vNormalInt, 1));
END_FOR
vTest2.ExecTime := LTIME() - vTest2.OldTime;

//------------CALCULATION C -------------------
vTest3.OldTime := LTIME();
FOR i:= 0 TO cRepeatCalcTimes DO
	setBitTovalue_bitmask(vNormalInt2, 2, checkBit_bitmask(vNormalInt2, 0) AND checkBit_bitmask(vNormalInt2, 1));
END_FOR
vTest3.ExecTime := LTIME() - vTest3.OldTime;


//------------CATCH RESULTS---------------------
vTest1.Results[vRunsCompleted] := vTest1.ExecTime;
vTest2.Results[vRunsCompleted] := vTest2.ExecTime;
vTest3.Results[vRunsCompleted] := vTest3.ExecTime;
              
END_ACTION
END_PROGRAM

PROGRAM x10_2_BitSet
  VAR CONSTANT
    cNrRuns : USINT(0..9) := 5;
    cRepeatCalcTimes : UDINT := 1000000;  (* 1 Million times *)
  END_VAR
  VAR_INPUT
    vStart : BOOL := FALSE;
  END_VAR
  VAR
    vDone : BOOL := FALSE;
    vRunsCompleted : USINT := 0;
    vStartTime : LTIME;
    vTotalTime : LTIME;
    vTest1 : dtSpeedTest;
    vTest2 : dtSpeedTest;
    vTest3 : dtSpeedTest;
    i : UDINT;
    vCodesysBits : dtBitStruct;  (* Test vars *)
    vNormalInt : UINT := 16#0;
    vNormalInt2 : UINT := 16#0;
    vNormalInt3 : UINT := 16#0;
    vResult1 : BOOL;
    vResult2 : BOOL;
    vResult3 : BOOL;
  END_VAR

            (*Runs once on event's rising edge*)
vDone 		:= FALSE;
vStartTime 	:= LTIME();

FOR vRunsCompleted:=0 TO cNrRuns DO
	Measure();
END_FOR

vTotalTime := LTIME() - vStartTime;

vTest1.Desc				:= 'Time to set bit 3, 1 Million times in codesys bit struct';
vTest1.AverageExecTime 	:= calcAvg(vTest1.Results);
vTest2.Desc				:= 'Time to set bit 3, 1 Million times in normal integer using . notation';
vTest2.AverageExecTime 	:= calcAvg(vTest2.Results);
vTest3.Desc				:= 'Time to set bit 3, 1 Million times in normal integer using bit masking';
vTest3.AverageExecTime 	:= calcAvg(vTest3.Results);
	
vDone := TRUE;
vStart:= FALSE;

          

ACTION Measure:
                //------------CALCULATION A -------------------
vTest1.OldTime := LTIME();
FOR i:= 0 TO cRepeatCalcTimes DO
	setBit_bitStruct(vCodesysBits, 2);
END_FOR
vTest1.ExecTime := LTIME() - vTest1.OldTime;

//------------CALCULATION B -------------------
vTest2.OldTime := LTIME();
FOR i:= 0 TO cRepeatCalcTimes DO
	setBit_dotNot(vNormalInt, 2);
END_FOR
vTest2.ExecTime := LTIME() - vTest2.OldTime;

//------------CALCULATION C -------------------
vTest3.OldTime := LTIME();
FOR i:= 0 TO cRepeatCalcTimes DO
	setBit_bitmask(vNormalInt2, 2);
END_FOR
vTest3.ExecTime := LTIME() - vTest3.OldTime;

//------------CATCH RESULTS---------------------
vTest1.Results[vRunsCompleted] := vTest1.ExecTime;
vTest2.Results[vRunsCompleted] := vTest2.ExecTime;
vTest3.Results[vRunsCompleted] := vTest3.ExecTime;
              
END_ACTION
END_PROGRAM

FUNCTION checkBit_bitmask : BOOL
  VAR_INPUT
    bits : UINT;
    bitToCheck : USINT;
  END_VAR

            checkBit_bitmask := (bits AND SHL(1, bitToCheck)) <> 0;
          
END_FUNCTION

FUNCTION setBit_bitmask : BOOL
  VAR_IN_OUT
    bits : UINT;
  END_VAR
  VAR_INPUT
    bitToSet : USINT;
  END_VAR

            bits := bits OR SHL(UINT#1, bitToSet);
          
END_FUNCTION

FUNCTION clearBit_bitmask : BOOL
  VAR_IN_OUT
    bits : UINT;
  END_VAR
  VAR_INPUT
    bitToClear : USINT;
  END_VAR

            bits := bits AND NOT SHL(UINT#1, bitToClear-1);
          
END_FUNCTION

FUNCTION setBitToValue_bitmask : BOOL
  VAR_IN_OUT
    bits : UINT;
  END_VAR
  VAR_INPUT
    bitToSet : USINT;
    value : BOOL;
  END_VAR

            IF value THEN
	setBit_bitmask(bits, bitToSet);
ELSE
	clearBit_bitmask(bits, bitToSet);
END_IF
          
END_FUNCTION

FUNCTION setBit_dotNot : BOOL
  VAR_IN_OUT
    bits : UINT;
  END_VAR
  VAR_INPUT
    bitToSet : USINT;
  END_VAR

            CASE bitToSet OF
	0: bits.0 := TRUE;
	1: bits.1 := TRUE;
	2: bits.2 := TRUE;
	3: bits.3 := TRUE;
	4: bits.4 := TRUE;
	5: bits.5 := TRUE;
	6: bits.6 := TRUE;
	7: bits.7 := TRUE;
	8: bits.8 := TRUE;
	9: bits.9 := TRUE;
	10: bits.10 := TRUE;
	11: bits.11 := TRUE;
	12: bits.12 := TRUE;
	13: bits.13 := TRUE;
	14: bits.14 := TRUE;
	15: bits.15 := TRUE;
END_CASE
          
END_FUNCTION

FUNCTION checkBit_dotNot : BOOL
  VAR_INPUT
    bits : UINT;
    bitToCheck : USINT;
  END_VAR

            CASE bitToCheck OF
	0: checkBit_dotNot := bits.0;
	1: checkBit_dotNot := bits.1;
	2: checkBit_dotNot := bits.2;
	3: checkBit_dotNot := bits.3;
	4: checkBit_dotNot := bits.4;
	5: checkBit_dotNot := bits.5;
	6: checkBit_dotNot := bits.6;
	7: checkBit_dotNot := bits.7;
	8: checkBit_dotNot := bits.8;
	9: checkBit_dotNot := bits.9;
	10: checkBit_dotNot := bits.10;
	11: checkBit_dotNot := bits.11;
	12: checkBit_dotNot := bits.12;
	13: checkBit_dotNot := bits.13;
	14: checkBit_dotNot := bits.14;
	15: checkBit_dotNot := bits.15;
END_CASE
          
END_FUNCTION

FUNCTION clearBit_dotNot : BOOL
  VAR_IN_OUT
    bits : UINT;
  END_VAR
  VAR_INPUT
    bitToClear : USINT;
  END_VAR

            CASE bitToClear OF
	0: bits.0 := FALSE;
	1: bits.1 := FALSE;
	2: bits.2 := FALSE;
	3: bits.3 := FALSE;
	4: bits.4 := FALSE;
	5: bits.5 := FALSE;
	6: bits.6 := FALSE;
	7: bits.7 := FALSE;
	8: bits.8 := FALSE;
	9: bits.9 := FALSE;
	10: bits.10 := FALSE;
	11: bits.11 := FALSE;
	12: bits.12 := FALSE;
	13: bits.13 := FALSE;
	14: bits.14 := FALSE;
	15: bits.15 := FALSE;
END_CASE
          
END_FUNCTION

FUNCTION checkBit_bitStruct : BOOL
  VAR_INPUT
    bits : dtBitStruct;
    bitToCheck : USINT;
  END_VAR

            CASE bitToCheck OF
	0: checkBit_bitStruct := bits.bit1;
	1: checkBit_bitStruct := bits.bit2;
	2: checkBit_bitStruct := bits.bit3;
	3: checkBit_bitStruct := bits.bit4;
	4: checkBit_bitStruct := bits.bit5;
	5: checkBit_bitStruct := bits.bit6;
	6: checkBit_bitStruct := bits.bit7;
	7: checkBit_bitStruct := bits.bit8;
	8: checkBit_bitStruct := bits.bit9;
	9: checkBit_bitStruct := bits.bit10;
	10: checkBit_bitStruct := bits.bit11;
	11: checkBit_bitStruct := bits.bit12;
	12: checkBit_bitStruct := bits.bit13;
	13: checkBit_bitStruct := bits.bit14;
	14: checkBit_bitStruct := bits.bit15;
	15: checkBit_bitStruct := bits.bit16;
END_CASE
          
END_FUNCTION

FUNCTION clearBit_bitStruct : BOOL
  VAR_IN_OUT
    bits : dtBitStruct;
  END_VAR
  VAR_INPUT
    bitToClear : USINT;
  END_VAR

            CASE bitToClear OF
	0: bits.bit1 := FALSE;
	1: bits.bit2 := FALSE;
	2: bits.bit3 := FALSE;
	3: bits.bit4 := FALSE;
	4: bits.bit5 := FALSE;
	5: bits.bit6 := FALSE;
	6: bits.bit7 := FALSE;
	7: bits.bit8 := FALSE;
	8: bits.bit9 := FALSE;
	9: bits.bit10 := FALSE;
	10: bits.bit11 := FALSE;
	11: bits.bit12 := FALSE;
	12: bits.bit13 := FALSE;
	13: bits.bit14 := FALSE;
	14: bits.bit15 := FALSE;
	15: bits.bit16 := FALSE;
END_CASE
          
END_FUNCTION

FUNCTION setBit_bitStruct : BOOL
  VAR_IN_OUT
    bits : dtBitStruct;
  END_VAR
  VAR_INPUT
    bitToSet : USINT;
  END_VAR

            CASE bitToSet OF
	0: bits.bit1 := TRUE;
	1: bits.bit2 := TRUE;
	2: bits.bit3 := TRUE;
	3: bits.bit4 := TRUE;
	4: bits.bit5 := TRUE;
	5: bits.bit6 := TRUE;
	6: bits.bit7 := TRUE;
	7: bits.bit8 := TRUE;
	8: bits.bit9 := TRUE;
	9: bits.bit10 := TRUE;
	10: bits.bit11 := TRUE;
	11: bits.bit12 := TRUE;
	12: bits.bit13 := TRUE;
	13: bits.bit14 := TRUE;
	14: bits.bit15 := TRUE;
	15: bits.bit16 := TRUE;
END_CASE
          
END_FUNCTION

FUNCTION setBitToValue_bitStruct : BOOL
  VAR_IN_OUT
    bits : dtBitStruct;
  END_VAR
  VAR_INPUT
    bitToSet : USINT;
    value : BOOL;
  END_VAR

            IF value THEN
	setBit_bitStruct(bits, bitToSet);
ELSE
	clearBit_bitStruct(bits, bitToSet);
END_IF
          
END_FUNCTION

FUNCTION setBitToValue_dotNot : BOOL
  VAR_IN_OUT
    bits : UINT;
  END_VAR
  VAR_INPUT
    bitToSet : USINT;
    value : BOOL;
  END_VAR

            IF value THEN
	setBit_dotNot(bits, bitToSet);
ELSE
	clearBit_dotNot(bits, bitToSet);
END_IF
          
END_FUNCTION

PROGRAM speedRunner
  VAR
    vTimeToRunTests : LTIME;
    vRunAll : BOOL;
  END_VAR

            (*Run tests one by one from the visu*)
(*or press the run all button*)
(*When run all is pressed, we must re trigger the event loop
also all these tests must run one by one
if run cyclically it messes up the total time*)
IF vRunAll THEN
	x01_ImpactOfDynamicArrays.vStart 	:= NOT x01_ImpactOfDynamicArrays.vDone;
	x02_ExecSpeedOfLanguageTypes.vStart := x01_ImpactOfDynamicArrays.vDone 		AND NOT x02_ExecSpeedOfLanguageTypes.vDone;
	x03_FloatingPointOperations.vStart 	:= x02_ExecSpeedOfLanguageTypes.vDone 	AND NOT x03_FloatingPointOperations.vDone;
	x04_FunctionOverhead.vStart 		:= x03_FloatingPointOperations.vDone 	AND NOT x04_FunctionOverhead.vDone;
	x05_SysMemLib.vStart 		:= x04_FunctionOverhead.vDone 			AND NOT x05_SysMemLib.vDone;
	x06_Combine2xByteToUint.vStart 				:= x05_SysMemLib.vDone 			AND NOT x06_Combine2xByteToUint.vDone;
	x07_StringOperations.vStart 		:= x06_Combine2xByteToUint.vDone 				AND NOT x07_StringOperations.vDone;
	x08_CheckingBools.vStart 			:= x07_StringOperations.vDone			AND NOT x08_CheckingBools.vDone;
	x09_CaseVsIfElsif.vStart 			:= x08_CheckingBools.vDone 				AND NOT x09_CaseVsIfElsif.vDone;
	x10_1_BitAccess.vStart 				:= x09_CaseVsIfElsif.vDone 				AND NOT x10_1_BitAccess.vDone;
	x10_2_BitSet.vStart 				:= x10_1_BitAccess.vDone 				AND NOT x10_2_BitSet.vDone;
	x10_3_BitMath.vStart 				:= x10_2_BitSet.vDone 					AND NOT x10_3_BitMath.vDone;
	x11_CalcInForLoppDecl.vStart 		:= x10_3_BitMath.vDone 					AND NOT x11_CalcInForLoppDecl.vDone;
	x12_BoolArrayToByteArray.vStart 	:= x11_CalcInForLoppDecl.vDone 			AND NOT x12_BoolArrayToByteArray.vDone;
	x13_ByteArrayToBool32.vStart 		:= x12_BoolArrayToByteArray.vDone 		AND NOT x13_ByteArrayToBool32.vDone;
END_IF

vTimeToRunTests :=  x01_ImpactOfDynamicArrays.vTotalTime + x02_ExecSpeedOfLanguageTypes.vTotalTime
					+ x03_FloatingPointOperations.vTotalTime + x04_FunctionOverhead.vTotalTime
					+ x05_SysMemLib.vTotalTime + x06_Combine2xByteToUint.vTotalTime
					+ x07_StringOperations.vTotalTime + x08_CheckingBools.vTotalTime
					+ x09_CaseVsIfElsif.vTotalTime + x10_1_BitAccess.vTotalTime
					+ x10_2_BitSet.vTotalTime + x10_3_BitMath.vTotalTime + x11_CalcInForLoppDecl.vTotalTime
					+ x12_BoolArrayToByteArray.vTotalTime + x13_ByteArrayToBool32.vTotalTime;
					


          
END_PROGRAM

FUNCTION calcMIPS : REAL
  VAR
    vMIPSOldTime : LTIME;
    i : DINT;
    vTestInt : UDINT;
    vMIPSExecTime : LTIME;
  END_VAR

            (*Calculate MIPS*)
vMIPSOldTime := LTIME();
FOR i:=1 TO 1000000 DO
	vTestInt := vTestInt + 1;
END_FOR
vMIPSExecTime := LTIME() - vMIPSOldTime;

(*Take a ratio of how long it took to add 1 milion integers, against 1 second, then divide by a milion to get MIPS(milion of integer additions per sec*)
calcMIPS := (vTestInt *  (1000000000.0 / LTIME_TO_REAL(vMIPSExecTime))) / 1000000.0;
          
END_FUNCTION

FUNCTION calcFLOPS : REAL
  VAR
    vFLOPSOldTime : LTIME;
    vTestReal : REAL;
    vFLOPSExecTime : LTIME;
    vMIPSAsReal : REAL;
    i : DINT;
  END_VAR

            (*Calculate FLOPS*)
vFLOPSOldTime := LTIME();
FOR i:=1 TO 1000000 DO
	vTestReal := vTestReal + 1.0;
END_FOR
vFLOPSExecTime := LTIME() - vFLOPSOldTime;

(*Take a ratio of how long it took to add 1 milion reals, against 1 second, then divide by a milion to get FLOPS(milion of floating point additions per sec*)
calcFLOPS := vTestReal *  (1000000000.0 / LTIME_TO_REAL(vFLOPSExecTime));
          
END_FUNCTION

PROGRAM x11_CalcInForLoppDecl
  VAR CONSTANT
    cNrRuns : USINT(0..9) := 5;
    cRepeatCalcTimes : UDINT := 10000;  (* 10 thousand times *)
  END_VAR
  VAR_INPUT
    vStart : BOOL := FALSE;
  END_VAR
  VAR
    vDone : BOOL := FALSE;
    vRunsCompleted : USINT := 0;
    vStartTime : LTIME;
    vTotalTime : LTIME;
    vTest1 : dtSpeedTest;
    vTest2 : dtSpeedTest;
    vTest3 : dtSpeedTest;
    i : UDINT;
    j : INT;
    vLongString : STRING(108) := '123456789123456789123456789123456789123456789123456789123456789123456789123456789123456789123456789123456789';  (* Test vars *)
    vResult : BYTE;
    vLenOfString : INT;
  END_VAR

            (*Runs once on event's rising edge*)
vDone 		:= FALSE;
vStartTime 	:= LTIME();

FOR vRunsCompleted:=0 TO cNrRuns DO
	Measure();
END_FOR

vTotalTime := LTIME() - vStartTime;

vTest1.Desc 			:= 'Time to iterate over bytes of a string[108] using known size, 10 thousand times';
vTest1.AverageExecTime 	:= calcAvg(vTest1.Results);
vTest2.Desc 			:= 'Time to iterate over bytes of a string[108] using calculation in declaration, 10 thousand times';
vTest2.AverageExecTime 	:= calcAvg(vTest2.Results);
vTest3.Desc 			:= 'Time to iterate over bytes of a STRING[108] using calculation outside OF the declaration, 10 thousand times';
vTest3.AverageExecTime 	:= calcAvg(vTest3.Results);
	
vDone := TRUE;
vStart:= FALSE;

          

ACTION Measure:
                //------------CALCULATION A -------------------
vTest1.OldTime := LTIME();
FOR i:= 0 TO cRepeatCalcTimes DO
	FOR j:= 0 TO 108 DO
		vResult := vLongString[j];
	END_FOR
END_FOR
vTest1.ExecTime := LTIME() - vTest1.OldTime;

//------------CALCULATION B -------------------
vTest2.OldTime := LTIME();
FOR i:= 0 TO cRepeatCalcTimes DO
	FOR j:= 0 TO LEN(vLongString) DO
		vResult := vLongString[j];
	END_FOR
END_FOR
vTest2.ExecTime := LTIME() - vTest2.OldTime;

//------------CALCULATION C -------------------
vTest3.OldTime := LTIME();
FOR i:= 0 TO cRepeatCalcTimes DO
	vLenOfString := LEN(vLongString);
	FOR j:= 0 TO vLenOfString DO
		vResult := vLongString[j];
	END_FOR
END_FOR
vTest3.ExecTime := LTIME() - vTest3.OldTime;

//------------CATCH RESULTS---------------------
vTest1.Results[vRunsCompleted] := vTest1.ExecTime;
vTest2.Results[vRunsCompleted] := vTest2.ExecTime;
vTest3.Results[vRunsCompleted] := vTest3.ExecTime;
              
END_ACTION
END_PROGRAM

PROGRAM x12_BoolArrayToByteArray
  VAR CONSTANT
    cNrRuns : USINT(0..9) := 5;
    cRepeatCalcTimes : UDINT := 1000000;  (* 1 Million times *)
  END_VAR
  VAR_INPUT
    vStart : BOOL := FALSE;
  END_VAR
  VAR
    vDone : BOOL := FALSE;
    vRunsCompleted : USINT := 0;
    vStartTime : LTIME;
    vTotalTime : LTIME;
    vTest1 : dtSpeedTest;
    vTest2 : dtSpeedTest;
    vTest3 : dtSpeedTest;
    vTest4 : dtSpeedTest;
    vTest5 : dtSpeedTest;
    vTest6 : dtSpeedTest;
    vTest7 : dtSpeedTest;
    i : UDINT;
    j : INT;
    vBoolArr : ARRAY[1..32] OF BOOL;  (* Test vars *)
    vBytes1 : ARRAY[1..4] OF USINT;
    vBytes2 : ARRAY[1..4] OF USINT;
    vBytes3 : ARRAY[1..4] OF USINT;
    vBytes4 : ARRAY[1..4] OF UINT;
    vBytes5 : ARRAY[1..4] OF UINT;
    vBytes6 : ARRAY[1..4] OF USINT;
    vBytes7 : ARRAY[1..4] OF USINT;
  END_VAR

            (*Runs once on event's rising edge*)
vDone 		:= FALSE;
vStartTime 	:= LTIME();

FOR vRunsCompleted:=0 TO cNrRuns DO
	Measure();
END_FOR

vTotalTime := LTIME() - vStartTime;

vTest1.Desc 			:= 'Time to pack bool array to 4 bytes, function, milion times';
vTest1.AverageExecTime 	:= calcAvg(vTest1.Results);
vTest2.Desc 			:= 'Time to pack bool array to 4 bytes, flat, milion times';
vTest2.AverageExecTime 	:= calcAvg(vTest2.Results);
vTest3.Desc 			:= 'Time TO pack bool array to 4 bytes, bitmask, milion times';
vTest3.AverageExecTime 	:= calcAvg(vTest3.Results);
vTest4.Desc 			:= 'Time to pack bool array to 4 bytes, bitmask function, milion times';
vTest4.AverageExecTime 	:= calcAvg(vTest4.Results);
vTest5.Desc 			:= 'Time TO pack bool array to 4 bytes, bitmask function in a loop, milion times';
vTest5.AverageExecTime 	:= calcAvg(vTest5.Results);
vTest6.Desc 			:= 'Time to pack bool array to 4 bytes, clear + bitmask, milion times';
vTest6.AverageExecTime 	:= calcAvg(vTest6.Results);
vTest7.Desc 			:= 'Time TO pack bool array to 4 bytes, clear + bitmask, function, milion times';
vTest7.AverageExecTime 	:= calcAvg(vTest7.Results);
	
vDone := TRUE;
vStart:= FALSE;

          

ACTION Measure:
                //------------CALCULATION A -------------------
vTest1.OldTime := LTIME();
FOR i:= 0 TO cRepeatCalcTimes DO
	vBytes1 := BOOLARR_TO_BYTES(vBoolArr);
END_FOR
vTest1.ExecTime := LTIME() - vTest1.OldTime;

//------------CALCULATION B -------------------
vTest2.OldTime := LTIME();
FOR i:= 0 TO cRepeatCalcTimes DO
	vBytes2[1].0 := vBoolArr[1];
	vBytes2[1].1 := vBoolArr[2];
	vBytes2[1].2 := vBoolArr[3];
	vBytes2[1].3 := vBoolArr[4];
	vBytes2[1].4 := vBoolArr[5];
	vBytes2[1].5 := vBoolArr[6];
	vBytes2[1].6 := vBoolArr[7];
	vBytes2[1].7 := vBoolArr[8];
	
	vBytes2[2].0 := vBoolArr[9];
	vBytes2[2].1 := vBoolArr[10];
	vBytes2[2].2 := vBoolArr[11];
	vBytes2[2].3 := vBoolArr[12];
	vBytes2[2].4 := vBoolArr[13];
	vBytes2[2].5 := vBoolArr[14];
	vBytes2[2].6 := vBoolArr[15];
	vBytes2[2].7 := vBoolArr[16];
	
	vBytes2[3].0 := vBoolArr[17];
	vBytes2[3].1 := vBoolArr[18];
	vBytes2[3].2 := vBoolArr[19];
	vBytes2[3].3 := vBoolArr[20];
	vBytes2[3].4 := vBoolArr[21];
	vBytes2[3].5 := vBoolArr[22];
	vBytes2[3].6 := vBoolArr[23];
	vBytes2[3].7 := vBoolArr[24];
	
	vBytes2[4].0 := vBoolArr[25];
	vBytes2[4].1 := vBoolArr[26];
	vBytes2[4].2 := vBoolArr[27];
	vBytes2[4].3 := vBoolArr[28];
	vBytes2[4].4 := vBoolArr[29];
	vBytes2[4].5 := vBoolArr[30];
	vBytes2[4].6 := vBoolArr[31];
	vBytes2[4].7 := vBoolArr[32];
END_FOR
vTest2.ExecTime := LTIME() - vTest2.OldTime;

//------------CALCULATION C -------------------
vTest3.OldTime := LTIME();
FOR i:= 0 TO cRepeatCalcTimes DO
	FOR j:=1 TO 4 DO
		vBytes3[j].0 := vBoolArr[1 + ((j-1) * 8)]; //1,9, 17, 25
		vBytes3[j].1 := vBoolArr[2 + ((j-1) * 8)];
		vBytes3[j].2 := vBoolArr[3 + ((j-1) * 8)];
		vBytes3[j].3 := vBoolArr[4 + ((j-1) * 8)];
		vBytes3[j].4 := vBoolArr[5 + ((j-1) * 8)];
		vBytes3[j].5 := vBoolArr[6 + ((j-1) * 8)]; //6, 14, 22, 30
		vBytes3[j].6 := vBoolArr[7 + ((j-1) * 8)]; //7, 15, 23, 31
		vBytes3[j].7 := vBoolArr[8 + ((j-1) * 8)]; //8, 16, 24, 32
	END_FOR
END_FOR
vTest3.ExecTime := LTIME() - vTest3.OldTime;

vTest4.OldTime := LTIME();
FOR i:= 0 TO cRepeatCalcTimes DO
	setBitToValue_bitmask(vBytes4[1], 1, vBoolArr[1]);
	setBitToValue_bitmask(vBytes4[1], 2 ,vBoolArr[2]);
	setBitToValue_bitmask(vBytes4[1], 3,vBoolArr[3]);
	setBitToValue_bitmask(vBytes4[1], 4,vBoolArr[4]);
	setBitToValue_bitmask(vBytes4[1], 5,vBoolArr[5]);
	setBitToValue_bitmask(vBytes4[1], 6,vBoolArr[6]);
	setBitToValue_bitmask(vBytes4[1], 7,vBoolArr[7]);
	setBitToValue_bitmask(vBytes4[1], 8,vBoolArr[8]);
	
	setBitToValue_bitmask(vBytes4[2], 1,vBoolArr[9]);
	setBitToValue_bitmask(vBytes4[2], 2,vBoolArr[10]);
	setBitToValue_bitmask(vBytes4[2], 3,vBoolArr[11]);
	setBitToValue_bitmask(vBytes4[2], 4,vBoolArr[12]);
	setBitToValue_bitmask(vBytes4[2], 5,vBoolArr[13]);
	setBitToValue_bitmask(vBytes4[2], 6,vBoolArr[14]);
	setBitToValue_bitmask(vBytes4[2], 7,vBoolArr[15]);
	setBitToValue_bitmask(vBytes4[2], 8,vBoolArr[16]);
	
	setBitToValue_bitmask(vBytes4[3], 1,vBoolArr[17]);
	setBitToValue_bitmask(vBytes4[3], 2,vBoolArr[18]);
	setBitToValue_bitmask(vBytes4[3], 3,vBoolArr[19]);
	setBitToValue_bitmask(vBytes4[3], 4,vBoolArr[20]);
	setBitToValue_bitmask(vBytes4[3], 5,vBoolArr[21]);
	setBitToValue_bitmask(vBytes4[3], 6,vBoolArr[22]);
	setBitToValue_bitmask(vBytes4[3], 7,vBoolArr[23]);
	setBitToValue_bitmask(vBytes4[3], 8,vBoolArr[24]);
	
	setBitToValue_bitmask(vBytes4[4], 1,vBoolArr[25]);
	setBitToValue_bitmask(vBytes4[4], 2,vBoolArr[26]);
	setBitToValue_bitmask(vBytes4[4], 3,vBoolArr[27]);
	setBitToValue_bitmask(vBytes4[4], 4,vBoolArr[28]);
	setBitToValue_bitmask(vBytes4[4], 5,vBoolArr[29]);
	setBitToValue_bitmask(vBytes4[4], 6,vBoolArr[30]);
	setBitToValue_bitmask(vBytes4[4], 7,vBoolArr[31]);
	setBitToValue_bitmask(vBytes4[4], 8,vBoolArr[32]);
END_FOR
vTest4.ExecTime := LTIME() - vTest4.OldTime;

vTest5.OldTime := LTIME();
FOR i:= 0 TO cRepeatCalcTimes DO
    FOR j:=1 TO 4 DO
        setBitToValue_bitmask(vBytes5[j], 1, vBoolArr[1 + ((j-1) * 8)]);
        setBitToValue_bitmask(vBytes5[j], 2, vBoolArr[2 + ((j-1) * 8)]);
        setBitToValue_bitmask(vBytes5[j], 3, vBoolArr[3 + ((j-1) * 8)]);
        setBitToValue_bitmask(vBytes5[j], 4, vBoolArr[4 + ((j-1) * 8)]);
        setBitToValue_bitmask(vBytes5[j], 5, vBoolArr[5 + ((j-1) * 8)]);
        setBitToValue_bitmask(vBytes5[j], 6, vBoolArr[6 + ((j-1) * 8)]);
        setBitToValue_bitmask(vBytes5[j], 7, vBoolArr[7 + ((j-1) * 8)]);
        setBitToValue_bitmask(vBytes5[j], 8, vBoolArr[8 + ((j-1) * 8)]);
    END_FOR
END_FOR
vTest5.ExecTime := LTIME() - vTest5.OldTime;


vTest6.OldTime := LTIME();
FOR i:= 0 TO cRepeatCalcTimes DO
    vBytes6[1] := 0;
    vBytes6[2] := 0;
    vBytes6[3] := 0;
    vBytes6[4] := 0;

	vBytes6[1] := vBytes6[1] OR SHL(BOOL_TO_USINT(vBoolArr[1]),0);
	vBytes6[1] := vBytes6[1] OR SHL(BOOL_TO_USINT(vBoolArr[2]),1);
	vBytes6[1] := vBytes6[1] OR SHL(BOOL_TO_USINT(vBoolArr[3]),2);
	vBytes6[1] := vBytes6[1] OR SHL(BOOL_TO_USINT(vBoolArr[4]),3);
	vBytes6[1] := vBytes6[1] OR SHL(BOOL_TO_USINT(vBoolArr[5]),4);
	vBytes6[1] := vBytes6[1] OR SHL(BOOL_TO_USINT(vBoolArr[6]),5);
	vBytes6[1] := vBytes6[1] OR SHL(BOOL_TO_USINT(vBoolArr[7]),6);
	vBytes6[1] := vBytes6[1] OR SHL(BOOL_TO_USINT(vBoolArr[8]),7);
	
	vBytes6[2] := vBytes6[2] OR SHL(BOOL_TO_USINT(vBoolArr[9]) ,0);
	vBytes6[2] := vBytes6[2] OR SHL(BOOL_TO_USINT(vBoolArr[10]),1);
	vBytes6[2] := vBytes6[2] OR SHL(BOOL_TO_USINT(vBoolArr[11]),2);
	vBytes6[2] := vBytes6[2] OR SHL(BOOL_TO_USINT(vBoolArr[12]),3);
	vBytes6[2] := vBytes6[2] OR SHL(BOOL_TO_USINT(vBoolArr[13]),4);
	vBytes6[2] := vBytes6[2] OR SHL(BOOL_TO_USINT(vBoolArr[14]),5);
	vBytes6[2] := vBytes6[2] OR SHL(BOOL_TO_USINT(vBoolArr[15]),6);
	vBytes6[2] := vBytes6[2] OR SHL(BOOL_TO_USINT(vBoolArr[16]),7);
	
	vBytes6[3] := vBytes6[3] OR SHL(BOOL_TO_USINT(vBoolArr[17]),0);
	vBytes6[3] := vBytes6[3] OR SHL(BOOL_TO_USINT(vBoolArr[18]),1);
	vBytes6[3] := vBytes6[3] OR SHL(BOOL_TO_USINT(vBoolArr[19]),2);
	vBytes6[3] := vBytes6[3] OR SHL(BOOL_TO_USINT(vBoolArr[20]),3);
	vBytes6[3] := vBytes6[3] OR SHL(BOOL_TO_USINT(vBoolArr[21]),4);
	vBytes6[3] := vBytes6[3] OR SHL(BOOL_TO_USINT(vBoolArr[22]),5);
	vBytes6[3] := vBytes6[3] OR SHL(BOOL_TO_USINT(vBoolArr[23]),6);
	vBytes6[3] := vBytes6[3] OR SHL(BOOL_TO_USINT(vBoolArr[24]),7);
	
	vBytes6[4] := vBytes6[4] OR SHL(BOOL_TO_USINT(vBoolArr[25]),0);
	vBytes6[4] := vBytes6[4] OR SHL(BOOL_TO_USINT(vBoolArr[26]),1);
	vBytes6[4] := vBytes6[4] OR SHL(BOOL_TO_USINT(vBoolArr[27]),2);
	vBytes6[4] := vBytes6[4] OR SHL(BOOL_TO_USINT(vBoolArr[28]),3);
	vBytes6[4] := vBytes6[4] OR SHL(BOOL_TO_USINT(vBoolArr[29]),4);
	vBytes6[4] := vBytes6[4] OR SHL(BOOL_TO_USINT(vBoolArr[30]),5);
	vBytes6[4] := vBytes6[4] OR SHL(BOOL_TO_USINT(vBoolArr[31]),6);
	vBytes6[4] := vBytes6[4] OR SHL(BOOL_TO_USINT(vBoolArr[32]),7);
END_FOR
vTest6.ExecTime := LTIME() - vTest6.OldTime;

vTest7.OldTime := LTIME();
FOR i:= 0 TO cRepeatCalcTimes DO
	vBytes7 := BOOLARR_TO_BYTES2(vBoolArr);
END_FOR
vTest7.ExecTime := LTIME() - vTest7.OldTime;

//------------CATCH RESULTS---------------------
vTest1.Results[vRunsCompleted] := vTest1.ExecTime;
vTest2.Results[vRunsCompleted] := vTest2.ExecTime;
vTest3.Results[vRunsCompleted] := vTest3.ExecTime;
vTest4.Results[vRunsCompleted] := vTest4.ExecTime;
vTest5.Results[vRunsCompleted] := vTest5.ExecTime;
vTest6.Results[vRunsCompleted] := vTest6.ExecTime;
vTest7.Results[vRunsCompleted] := vTest7.ExecTime;
              
END_ACTION
END_PROGRAM

FUNCTION BOOLARR_TO_BYTES : ARRAY[1..4] OF USINT
  VAR_IN_OUT
    Data : ARRAY[1..32] OF BOOL;
  END_VAR

            BOOLARR_TO_BYTES[1].0 := Data[1];
BOOLARR_TO_BYTES[1].1 := Data[2];
BOOLARR_TO_BYTES[1].2 := Data[3];
BOOLARR_TO_BYTES[1].3 := Data[4];
BOOLARR_TO_BYTES[1].4 := Data[5];
BOOLARR_TO_BYTES[1].5 := Data[6];
BOOLARR_TO_BYTES[1].6 := Data[7];
BOOLARR_TO_BYTES[1].7 := Data[8];

BOOLARR_TO_BYTES[2].0 := Data[9];
BOOLARR_TO_BYTES[2].1 := Data[10];
BOOLARR_TO_BYTES[2].2 := Data[11];
BOOLARR_TO_BYTES[2].3 := Data[12];
BOOLARR_TO_BYTES[2].4 := Data[13];
BOOLARR_TO_BYTES[2].5 := Data[14];
BOOLARR_TO_BYTES[2].6 := Data[15];
BOOLARR_TO_BYTES[2].7 := Data[16];

BOOLARR_TO_BYTES[3].0 := Data[17];
BOOLARR_TO_BYTES[3].1 := Data[18];
BOOLARR_TO_BYTES[3].2 := Data[19];
BOOLARR_TO_BYTES[3].3 := Data[20];
BOOLARR_TO_BYTES[3].4 := Data[21];
BOOLARR_TO_BYTES[3].5 := Data[22];
BOOLARR_TO_BYTES[3].6 := Data[23];
BOOLARR_TO_BYTES[3].7 := Data[24];

BOOLARR_TO_BYTES[4].0 := Data[25];
BOOLARR_TO_BYTES[4].1 := Data[26];
BOOLARR_TO_BYTES[4].2 := Data[27];
BOOLARR_TO_BYTES[4].3 := Data[28];
BOOLARR_TO_BYTES[4].4 := Data[29];
BOOLARR_TO_BYTES[4].5 := Data[30];
BOOLARR_TO_BYTES[4].6 := Data[31];
BOOLARR_TO_BYTES[4].7 := Data[32];
          
END_FUNCTION

FUNCTION BOOLARR_TO_BYTES2 : ARRAY[1..4] OF USINT
  VAR_IN_OUT
    Data : ARRAY[1..32] OF BOOL;
  END_VAR

            BOOLARR_TO_BYTES2[1] := BOOLARR_TO_BYTES2[1] OR SHL(BOOL_TO_USINT(Data[1]),0);
BOOLARR_TO_BYTES2[1] := BOOLARR_TO_BYTES2[1] OR SHL(BOOL_TO_USINT(Data[2]),1);
BOOLARR_TO_BYTES2[1] := BOOLARR_TO_BYTES2[1] OR SHL(BOOL_TO_USINT(Data[3]),2);
BOOLARR_TO_BYTES2[1] := BOOLARR_TO_BYTES2[1] OR SHL(BOOL_TO_USINT(Data[4]),3);
BOOLARR_TO_BYTES2[1] := BOOLARR_TO_BYTES2[1] OR SHL(BOOL_TO_USINT(Data[5]),4);
BOOLARR_TO_BYTES2[1] := BOOLARR_TO_BYTES2[1] OR SHL(BOOL_TO_USINT(Data[6]),5);
BOOLARR_TO_BYTES2[1] := BOOLARR_TO_BYTES2[1] OR SHL(BOOL_TO_USINT(Data[7]),6);
BOOLARR_TO_BYTES2[1] := BOOLARR_TO_BYTES2[1] OR SHL(BOOL_TO_USINT(Data[8]),7);
	
BOOLARR_TO_BYTES2[2] := BOOLARR_TO_BYTES2[2] OR SHL(BOOL_TO_USINT(Data[9]) ,0);
BOOLARR_TO_BYTES2[2] := BOOLARR_TO_BYTES2[2] OR SHL(BOOL_TO_USINT(Data[10]),1);
BOOLARR_TO_BYTES2[2] := BOOLARR_TO_BYTES2[2] OR SHL(BOOL_TO_USINT(Data[11]),2);
BOOLARR_TO_BYTES2[2] := BOOLARR_TO_BYTES2[2] OR SHL(BOOL_TO_USINT(Data[12]),3);
BOOLARR_TO_BYTES2[2] := BOOLARR_TO_BYTES2[2] OR SHL(BOOL_TO_USINT(Data[13]),4);
BOOLARR_TO_BYTES2[2] := BOOLARR_TO_BYTES2[2] OR SHL(BOOL_TO_USINT(Data[14]),5);
BOOLARR_TO_BYTES2[2] := BOOLARR_TO_BYTES2[2] OR SHL(BOOL_TO_USINT(Data[15]),6);
BOOLARR_TO_BYTES2[2] := BOOLARR_TO_BYTES2[2] OR SHL(BOOL_TO_USINT(Data[16]),7);
	
BOOLARR_TO_BYTES2[3] := BOOLARR_TO_BYTES2[3] OR SHL(BOOL_TO_USINT(Data[17]),0);
BOOLARR_TO_BYTES2[3] := BOOLARR_TO_BYTES2[3] OR SHL(BOOL_TO_USINT(Data[18]),1);
BOOLARR_TO_BYTES2[3] := BOOLARR_TO_BYTES2[3] OR SHL(BOOL_TO_USINT(Data[19]),2);
BOOLARR_TO_BYTES2[3] := BOOLARR_TO_BYTES2[3] OR SHL(BOOL_TO_USINT(Data[20]),3);
BOOLARR_TO_BYTES2[3] := BOOLARR_TO_BYTES2[3] OR SHL(BOOL_TO_USINT(Data[21]),4);
BOOLARR_TO_BYTES2[3] := BOOLARR_TO_BYTES2[3] OR SHL(BOOL_TO_USINT(Data[22]),5);
BOOLARR_TO_BYTES2[3] := BOOLARR_TO_BYTES2[3] OR SHL(BOOL_TO_USINT(Data[23]),6);
BOOLARR_TO_BYTES2[3] := BOOLARR_TO_BYTES2[3] OR SHL(BOOL_TO_USINT(Data[24]),7);
	
BOOLARR_TO_BYTES2[4] := BOOLARR_TO_BYTES2[4] OR SHL(BOOL_TO_USINT(Data[25]),0);
BOOLARR_TO_BYTES2[4] := BOOLARR_TO_BYTES2[4] OR SHL(BOOL_TO_USINT(Data[26]),1);
BOOLARR_TO_BYTES2[4] := BOOLARR_TO_BYTES2[4] OR SHL(BOOL_TO_USINT(Data[27]),2);
BOOLARR_TO_BYTES2[4] := BOOLARR_TO_BYTES2[4] OR SHL(BOOL_TO_USINT(Data[28]),3);
BOOLARR_TO_BYTES2[4] := BOOLARR_TO_BYTES2[4] OR SHL(BOOL_TO_USINT(Data[29]),4);
BOOLARR_TO_BYTES2[4] := BOOLARR_TO_BYTES2[4] OR SHL(BOOL_TO_USINT(Data[30]),5);
BOOLARR_TO_BYTES2[4] := BOOLARR_TO_BYTES2[4] OR SHL(BOOL_TO_USINT(Data[31]),6);
BOOLARR_TO_BYTES2[4] := BOOLARR_TO_BYTES2[4] OR SHL(BOOL_TO_USINT(Data[32]),7);
          
END_FUNCTION

PROGRAM x13_ByteArrayToBool32
  VAR CONSTANT
    cNrRuns : USINT(0..9) := 5;
    cRepeatCalcTimes : UDINT := 1000000;  (* 1 Million times *)
  END_VAR
  VAR_INPUT
    vStart : BOOL := FALSE;
  END_VAR
  VAR
    vDone : BOOL := FALSE;
    vRunsCompleted : USINT := 0;
    vStartTime : LTIME;
    vTotalTime : LTIME;
    vTest1 : dtSpeedTest;
    vTest2 : dtSpeedTest;
    vTest3 : dtSpeedTest;
    vTest4 : dtSpeedTest;
    i : UDINT;
    j : INT;
    vBoolArr1 : ARRAY[1..32] OF BOOL;  (* Test vars *)
    vBoolArr2 : ARRAY[1..32] OF BOOL;
    vBoolArr3 : ARRAY[1..32] OF BOOL;
    vBoolArr4 : ARRAY[1..32] OF BOOL;
    vBytes : ARRAY[1..4] OF USINT := [16#FF, 16#85, 16#0, 16#AB];
  END_VAR

            (*Runs once on event's rising edge*)
vDone 		:= FALSE;
vStartTime 	:= LTIME();

FOR vRunsCompleted:=0 TO cNrRuns DO
	Measure();
END_FOR

vTotalTime := LTIME() - vStartTime;

vTest1.Desc 			:= 'Time to upack 4 bytes to bool array, function, milion times';
vTest1.AverageExecTime 	:= calcAvg(vTest1.Results);
vTest2.Desc 			:= 'Time to upack 4 bytes to bool array, flat, milion times, milion times';
vTest2.AverageExecTime 	:= calcAvg(vTest2.Results);
vTest3.Desc 			:= 'Time to upack 4 bytes to bool array, bitmask function, milion times, milion times';
vTest3.AverageExecTime 	:= calcAvg(vTest3.Results);
vTest4.Desc 			:= 'Time to upack 4 bytes to bool array, bitmask, milion times, milion times';
vTest4.AverageExecTime 	:= calcAvg(vTest4.Results);

vDone := TRUE;
vStart:= FALSE;

          

ACTION Measure:
                //------------CALCULATION A -------------------
vTest1.OldTime := LTIME();
FOR i:= 0 TO cRepeatCalcTimes DO
	vBoolArr1 := UnpackBytesToBool32(vBytes);
END_FOR
vTest1.ExecTime := LTIME() - vTest1.OldTime;

//------------CALCULATION B -------------------
vTest2.OldTime := LTIME();
FOR i:= 0 TO cRepeatCalcTimes DO
	vBoolArr2[1] := vBytes[1].0;
	vBoolArr2[2] := vBytes[1].1;
	vBoolArr2[3] := vBytes[1].2;
	vBoolArr2[4] := vBytes[1].3;
	vBoolArr2[5] := vBytes[1].4;
	vBoolArr2[6] := vBytes[1].5;
	vBoolArr2[7] := vBytes[1].6;
	vBoolArr2[8] := vBytes[1].7;
	
	vBoolArr2[9] :=  vBytes[2].0;
	vBoolArr2[10] := vBytes[2].1;
	vBoolArr2[11] := vBytes[2].2;
	vBoolArr2[12] := vBytes[2].3;
	vBoolArr2[13] := vBytes[2].4;
	vBoolArr2[14] := vBytes[2].5;
	vBoolArr2[15] := vBytes[2].6;
	vBoolArr2[16] := vBytes[2].7;
	
	vBoolArr2[17] := vBytes[3].0;
	vBoolArr2[18] := vBytes[3].1;
	vBoolArr2[19] := vBytes[3].2;
	vBoolArr2[20] := vBytes[3].3;
	vBoolArr2[21] := vBytes[3].4;
	vBoolArr2[22] := vBytes[3].5;
	vBoolArr2[23] := vBytes[3].6;
	vBoolArr2[24] := vBytes[3].7;
	
	vBoolArr2[25] := vBytes[4].0;
	vBoolArr2[26] := vBytes[4].1;
	vBoolArr2[27] := vBytes[4].2;
	vBoolArr2[28] := vBytes[4].3;
	vBoolArr2[29] := vBytes[4].4;
	vBoolArr2[30] := vBytes[4].5;
	vBoolArr2[31] := vBytes[4].6;
	vBoolArr2[32] := vBytes[4].7;

END_FOR
vTest2.ExecTime := LTIME() - vTest2.OldTime;

//------------CALCULATION C -------------------
vTest3.OldTime := LTIME();
FOR i:= 0 TO cRepeatCalcTimes DO
	vBoolArr3 := UnpackBytesToBool32_2(vBytes);
END_FOR
vTest3.ExecTime := LTIME() - vTest3.OldTime;

vTest4.OldTime := LTIME();
FOR i:= 0 TO cRepeatCalcTimes DO
	vBoolArr4[1] := (vBytes[1] AND 1) <> 0;
	vBoolArr4[2] := (vBytes[1] AND 2) <> 0;
	vBoolArr4[3] := (vBytes[1] AND 4) <> 0;
	vBoolArr4[4] := (vBytes[1] AND 8) <> 0;
	vBoolArr4[5] := (vBytes[1] AND 16) <> 0;
	vBoolArr4[6] := (vBytes[1] AND 32) <> 0;
	vBoolArr4[7] := (vBytes[1] AND 64) <> 0;
	vBoolArr4[8] := (vBytes[1] AND 128) <> 0;
	
	vBoolArr4[9] := (vBytes[2] AND  1) <> 0;
	vBoolArr4[10] := (vBytes[2] AND 2) <> 0;
	vBoolArr4[11] := (vBytes[2] AND 4) <> 0;
	vBoolArr4[12] := (vBytes[2] AND 8) <> 0;
	vBoolArr4[13] := (vBytes[2] AND 16) <> 0;
	vBoolArr4[14] := (vBytes[2] AND 32) <> 0;
	vBoolArr4[15] := (vBytes[2] AND 64) <> 0;
	vBoolArr4[16] := (vBytes[2] AND 128) <> 0;
	
	vBoolArr4[17] := (vBytes[3] AND 1) <> 0;
	vBoolArr4[18] := (vBytes[3] AND 2) <> 0;
	vBoolArr4[19] := (vBytes[3] AND 4) <> 0;
	vBoolArr4[20] := (vBytes[3] AND 8) <> 0;
	vBoolArr4[21] := (vBytes[3] AND 16) <> 0;
	vBoolArr4[22] := (vBytes[3] AND 32) <> 0;
	vBoolArr4[23] := (vBytes[3] AND 64) <> 0;
	vBoolArr4[24] := (vBytes[3] AND 128) <> 0;
	
	vBoolArr4[25] := (vBytes[4] AND 1) <> 0;
	vBoolArr4[26] := (vBytes[4] AND 2) <> 0;
	vBoolArr4[27] := (vBytes[4] AND 4) <> 0;
	vBoolArr4[28] := (vBytes[4] AND 8) <> 0;
	vBoolArr4[29] := (vBytes[4] AND 16) <> 0;
	vBoolArr4[30] := (vBytes[4] AND 32) <> 0;
	vBoolArr4[31] := (vBytes[4] AND 64) <> 0;
	vBoolArr4[32] := (vBytes[4] AND 128) <> 0;

END_FOR
vTest4.ExecTime := LTIME() - vTest4.OldTime;

//------------CATCH RESULTS---------------------
vTest1.Results[vRunsCompleted] := vTest1.ExecTime;
vTest2.Results[vRunsCompleted] := vTest2.ExecTime;
vTest3.Results[vRunsCompleted] := vTest3.ExecTime;
vTest4.Results[vRunsCompleted] := vTest4.ExecTime;
              
END_ACTION
END_PROGRAM

FUNCTION UnpackBytesToBool32 : ARRAY[1..32] OF BOOL
  VAR_IN_OUT
    Bytes : ARRAY[1..4] OF USINT;
  END_VAR

            UnpackBytesToBool32[1] := Bytes[1].0;
UnpackBytesToBool32[2] := Bytes[1].1;
UnpackBytesToBool32[3] := Bytes[1].2;
UnpackBytesToBool32[4] := Bytes[1].3;
UnpackBytesToBool32[5] := Bytes[1].4;
UnpackBytesToBool32[6] := Bytes[1].5;
UnpackBytesToBool32[7] := Bytes[1].6;
UnpackBytesToBool32[8] := Bytes[1].7;

UnpackBytesToBool32[9] := Bytes[2].0;
UnpackBytesToBool32[10] := Bytes[2].1;
UnpackBytesToBool32[11] := Bytes[2].2;
UnpackBytesToBool32[12] := Bytes[2].3;
UnpackBytesToBool32[13] := Bytes[2].4;
UnpackBytesToBool32[14] := Bytes[2].5;
UnpackBytesToBool32[15] := Bytes[2].6;
UnpackBytesToBool32[16] := Bytes[2].7;

UnpackBytesToBool32[17] := Bytes[3].0;
UnpackBytesToBool32[18] := Bytes[3].1;
UnpackBytesToBool32[19] := Bytes[3].2;
UnpackBytesToBool32[20] := Bytes[3].3;
UnpackBytesToBool32[21] := Bytes[3].4;
UnpackBytesToBool32[22] := Bytes[3].5;
UnpackBytesToBool32[23] := Bytes[3].6;
UnpackBytesToBool32[24] := Bytes[3].7;

UnpackBytesToBool32[25] := Bytes[4].0;
UnpackBytesToBool32[26] := Bytes[4].1;
UnpackBytesToBool32[27] := Bytes[4].2;
UnpackBytesToBool32[28] := Bytes[4].3;
UnpackBytesToBool32[29] := Bytes[4].4;
UnpackBytesToBool32[30] := Bytes[4].5;
UnpackBytesToBool32[31] := Bytes[4].6;
UnpackBytesToBool32[32] := Bytes[4].7;

          
END_FUNCTION

FUNCTION UnpackBytesToBool32_2 : ARRAY[1..32] OF BOOL
  VAR_IN_OUT
    Bytes : ARRAY[1..4] OF USINT;
  END_VAR

            UnpackBytesToBool32_2[1] := (Bytes[1] AND 1) <> 0;
UnpackBytesToBool32_2[2] := (Bytes[1] AND 2) <> 0;
UnpackBytesToBool32_2[3] := (Bytes[1] AND 4) <> 0;
UnpackBytesToBool32_2[4] := (Bytes[1] AND 8) <> 0;
UnpackBytesToBool32_2[5] := (Bytes[1] AND 16) <> 0;
UnpackBytesToBool32_2[6] := (Bytes[1] AND 32) <> 0;
UnpackBytesToBool32_2[7] := (Bytes[1] AND 64) <> 0;
UnpackBytesToBool32_2[8] := (Bytes[1] AND 128) <> 0;

UnpackBytesToBool32_2[9] :=  (Bytes[2] AND 1) <> 0;;
UnpackBytesToBool32_2[10] := (Bytes[2] AND 2) <> 0;
UnpackBytesToBool32_2[11] := (Bytes[2] AND 4) <> 0;
UnpackBytesToBool32_2[12] := (Bytes[2] AND 8) <> 0;
UnpackBytesToBool32_2[13] := (Bytes[2] AND 16) <> 0;
UnpackBytesToBool32_2[14] := (Bytes[2] AND 32) <> 0;
UnpackBytesToBool32_2[15] := (Bytes[2] AND 64) <> 0;
UnpackBytesToBool32_2[16] := (Bytes[2] AND 128) <> 0;

UnpackBytesToBool32_2[17] := (Bytes[3] AND 1) <> 0;
UnpackBytesToBool32_2[18] := (Bytes[3] AND 2) <> 0;
UnpackBytesToBool32_2[19] := (Bytes[3] AND 4) <> 0;
UnpackBytesToBool32_2[20] := (Bytes[3] AND 8) <> 0;
UnpackBytesToBool32_2[21] := (Bytes[3] AND 16) <> 0;
UnpackBytesToBool32_2[22] := (Bytes[3] AND 32) <> 0;
UnpackBytesToBool32_2[23] := (Bytes[3] AND 64) <> 0;
UnpackBytesToBool32_2[24] := (Bytes[3] AND 128) <> 0;

UnpackBytesToBool32_2[25] := (Bytes[4] AND 1) <> 0;
UnpackBytesToBool32_2[26] := (Bytes[4] AND 2) <> 0;
UnpackBytesToBool32_2[27] := (Bytes[4] AND 4) <> 0;
UnpackBytesToBool32_2[28] := (Bytes[4] AND 8) <> 0;
UnpackBytesToBool32_2[29] := (Bytes[4] AND 16) <> 0;
UnpackBytesToBool32_2[30] := (Bytes[4] AND 32) <> 0;
UnpackBytesToBool32_2[31] := (Bytes[4] AND 64) <> 0;
UnpackBytesToBool32_2[32] := (Bytes[4] AND 128) <> 0;

          
END_FUNCTION

PROGRAM x00_CalcMIPS_FLOPS
  VAR
    vStart : BOOL;
    vDone : BOOL;
    vMIPS : REAL;
    vFLOPS : REAL;
    vkFLOPS : REAL;
    vMFLOPS : REAL;
    vGFLOPS : REAL;
  END_VAR

            vDone := FALSE;
(*Calculate MIPS and FLOPS of this machine
	PS: These calcs are not 100% accurate but more to compare machine to machine*)
(*
	System spec:
	- OS Name	Microsoft Windows 10 Home	
	- Version	10.0.19044 Build 19044	
	- OS Manufacturer	Microsoft Corporation	
	- System Manufacturer	SAMSUNG ELECTRONICS CO., LTD.	
	- System Model	3570R/370R/470R/450R/510R/4450RV	
	- System Type	x64-based PC	
	- Processor	Intel(R) Core(TM) i5-3210M CPU @ 2.50GHz, 2501 Mhz, 2 Core(s), 4 Logical Processor(s)	
	- Installed Physical Memory (RAM)	8,00 GB	
	- Total Physical Memory	7,89 GB	
	- Available Physical Memory	3,80 GB	
	- Total Virtual Memory	9,75 GB	
	- Available Virtual Memory	5,66 GB	
	
	MIPS 	-> 407
	FLOPS 	-> 3.32e+08
	kFLOPS 	-> 3.32e+05
	MFLOPS 	-> 332
	GFLOPS 	-> 0.332
*)
vMIPS 	:= calcMIPS();
vFLOPS	:= calcFLOPS();
vkFLOPS := vFLOPS / 1000.0;
vMFLOPS := vFLOPS / 1000000.0;
vGFLOPS := vFLOPS / (1000.0 * 1000000.0);

vDone := TRUE;
          
END_PROGRAM

FUNCTION calcAvgFixed : LTIME
  VAR_IN_OUT
    Results : ARRAY[0..9] OF LTIME;
  END_VAR
  VAR
    i : USINT;
  END_VAR

            FOR i:=0 TO 9 DO
	IF Results[i] = LTIME#0S THEN
		EXIT;
	END_IF
	calcAvgFixed := calcAvgFixed + Results[i];
END_FOR
calcAvgFixed := calcAvgFixed / MAX(1,i);
RETURN;
          
END_FUNCTION

FUNCTION addTwoIntsCFC : INT
  VAR_INPUT
    int1 : INT;
    int2 : INT;
  END_VAR
  VAR  (* added by the conversion: wires and edge detectors of the diagram *)
    _ADD2_OUT : ANY;
  END_VAR

(* CFC diagram, written out as Structured Text *)
addTwoIntsCFC := _ADD2_OUT;
_ADD2_OUT := int1 + int2;
END_FUNCTION

CONFIGURATION CODESYS_Control_Win_V3_x64
  RESOURCE Application ON PLC
    TASK SpdRnnr(INTERVAL := T#200ms, PRIORITY := 16);
    TASK VISU_TASK(INTERVAL := T#200ms, PRIORITY := 31);
    TASK x01(SINGLE := x01_ImpactOfDynamicArrays.vStart, PRIORITY := 1);
    TASK x02(SINGLE := x02_ExecSpeedOfLanguageTypes.vStart, PRIORITY := 1);
    TASK x04(SINGLE := x04_FunctionOverhead.vStart, PRIORITY := 1);
    TASK x05(SINGLE := x05_SysMemLib.vStart, PRIORITY := 1);
    TASK x06(SINGLE := x06_Combine2xByteToUint.vStart, PRIORITY := 1);
    TASK x07(SINGLE := x07_StringOperations.vStart, PRIORITY := 1);
    TASK x08(SINGLE := x08_CheckingBools.vStart, PRIORITY := 1);
    TASK x09(SINGLE := x09_CaseVsIfElsif.vStart, PRIORITY := 1);
    TASK x10_1(SINGLE := x10_1_BitAccess.vStart, PRIORITY := 1);
    TASK x11(SINGLE := x11_CalcInForLoppDecl.vStart, PRIORITY := 1);
    TASK x03(SINGLE := x03_FloatingPointOperations.vStart, PRIORITY := 1);
    TASK x12(SINGLE := x12_BoolArrayToByteArray.vStart, PRIORITY := 1);
    TASK x13(SINGLE := x13_ByteArrayToBool32.vStart, PRIORITY := 1);
    TASK x10_2(SINGLE := x10_2_BitSet.vStart, PRIORITY := 1);
    TASK x10_3(SINGLE := x10_3_BitMath.vStart, PRIORITY := 1);
    TASK x00(SINGLE := x00_CalcMIPS_FLOPS.vStart, PRIORITY := 1);
    PROGRAM speedRunner WITH SpdRnnr : speedRunner;
    PROGRAM VisuElems.Visu_Prg WITH VISU_TASK : VisuElems.Visu_Prg;
    PROGRAM x01_ImpactOfDynamicArrays WITH x01 : x01_ImpactOfDynamicArrays;
    PROGRAM x02_ExecSpeedOfLanguageTypes WITH x02 : x02_ExecSpeedOfLanguageTypes;
    PROGRAM x04_FunctionOverhead WITH x04 : x04_FunctionOverhead;
    PROGRAM x05_SysMemLib WITH x05 : x05_SysMemLib;
    PROGRAM x06_Combine2xByteToUint WITH x06 : x06_Combine2xByteToUint;
    PROGRAM x07_StringOperations WITH x07 : x07_StringOperations;
    PROGRAM x08_CheckingBools WITH x08 : x08_CheckingBools;
    PROGRAM x09_CaseVsIfElsif WITH x09 : x09_CaseVsIfElsif;
    PROGRAM x10_1_BitAccess WITH x10_1 : x10_1_BitAccess;
    PROGRAM x11_CalcInForLoppDecl WITH x11 : x11_CalcInForLoppDecl;
    PROGRAM x03_FloatingPointOperations WITH x03 : x03_FloatingPointOperations;
    PROGRAM x12_BoolArrayToByteArray WITH x12 : x12_BoolArrayToByteArray;
    PROGRAM x13_ByteArrayToBool32 WITH x13 : x13_ByteArrayToBool32;
    PROGRAM x10_2_BitSet WITH x10_2 : x10_2_BitSet;
    PROGRAM x10_3_BitMath WITH x10_3 : x10_3_BitMath;
    PROGRAM x00_CalcMIPS_FLOPS WITH x00 : x00_CalcMIPS_FLOPS;
  END_RESOURCE
END_CONFIGURATION

CONFIGURATION CODESYS_Control_RTE_V3_x64
  RESOURCE Application ON PLC
    TASK x01(SINGLE := x01_ImpactOfDynamicArrays.vStart, PRIORITY := 1);
    TASK x04(SINGLE := x04_FunctionOverhead.vStart, PRIORITY := 1);
    TASK SpdRnnr(INTERVAL := T#200ms, PRIORITY := 16);
    TASK x06(SINGLE := x06_Combine2xByteToUint.vStart, PRIORITY := 1);
    TASK x02(SINGLE := x02_ExecSpeedOfLanguageTypes.vStart, PRIORITY := 1);
    TASK VISU_TASK(INTERVAL := T#200ms, PRIORITY := 31);
    TASK x07(SINGLE := x07_StringOperations.vStart, PRIORITY := 1);
    TASK x08(SINGLE := x08_CheckingBools.vStart, PRIORITY := 1);
    TASK x10_1(SINGLE := x10_1_BitAccess.vStart, PRIORITY := 1);
    TASK x09(SINGLE := x09_CaseVsIfElsif.vStart, PRIORITY := 1);
    TASK x05(SINGLE := x05_SysMemLib.vStart, PRIORITY := 1);
    TASK x12(SINGLE := x12_BoolArrayToByteArray.vStart, PRIORITY := 1);
    TASK x13(SINGLE := x13_ByteArrayToBool32.vStart, PRIORITY := 1);
    TASK x11(SINGLE := x11_CalcInForLoppDecl.vStart, PRIORITY := 1);
    TASK x03(SINGLE := x03_FloatingPointOperations.vStart, PRIORITY := 1);
    TASK x10_2(SINGLE := x10_2_BitSet.vStart, PRIORITY := 1);
    TASK x10_3(SINGLE := x10_3_BitMath.vStart, PRIORITY := 1);
    TASK x00(SINGLE := x00_CalcMIPS_FLOPS.vStart, PRIORITY := 1);
    PROGRAM x01_ImpactOfDynamicArrays WITH x01 : x01_ImpactOfDynamicArrays;
    PROGRAM x04_FunctionOverhead WITH x04 : x04_FunctionOverhead;
    PROGRAM speedRunner WITH SpdRnnr : speedRunner;
    PROGRAM x06_Combine2xByteToUint WITH x06 : x06_Combine2xByteToUint;
    PROGRAM x02_ExecSpeedOfLanguageTypes WITH x02 : x02_ExecSpeedOfLanguageTypes;
    PROGRAM VisuElems.Visu_Prg WITH VISU_TASK : VisuElems.Visu_Prg;
    PROGRAM x07_StringOperations WITH x07 : x07_StringOperations;
    PROGRAM x08_CheckingBools WITH x08 : x08_CheckingBools;
    PROGRAM x10_1_BitAccess WITH x10_1 : x10_1_BitAccess;
    PROGRAM x09_CaseVsIfElsif WITH x09 : x09_CaseVsIfElsif;
    PROGRAM x05_SysMemLib WITH x05 : x05_SysMemLib;
    PROGRAM x12_BoolArrayToByteArray WITH x12 : x12_BoolArrayToByteArray;
    PROGRAM x13_ByteArrayToBool32 WITH x13 : x13_ByteArrayToBool32;
    PROGRAM x11_CalcInForLoppDecl WITH x11 : x11_CalcInForLoppDecl;
    PROGRAM x03_FloatingPointOperations WITH x03 : x03_FloatingPointOperations;
    PROGRAM x10_2_BitSet WITH x10_2 : x10_2_BitSet;
    PROGRAM x10_3_BitMath WITH x10_3 : x10_3_BitMath;
    PROGRAM x00_CalcMIPS_FLOPS WITH x00 : x00_CalcMIPS_FLOPS;
  END_RESOURCE
END_CONFIGURATION
